(* IEC 61131-3 sources: daoli-st-library/DL_Motion (part 19) *)

(* ---- FB_DL_StringCutAlign.st ---- *)
(*==============================================================================
 * 组件名称 (Component)  : FB_DL_StringCutAlign
 * 所属子库 (Sublibrary) : DL_Motion
 * 当前版本 (Version)    : 1.0.0
 * 兼容性 (Platform)     : CODESYS 3.5 / TwinCAT 3 / 汇川 InoProShop / Machine Expert
 *                         仅依赖纯 IEC 61131-3 标准元素，零厂商方言
 * 功能描述 (Function)   : 串焊裁切对位：bCutCycle 上升沿锁存相机偏差 → 委托
 *                         FB_DL_LowPassFilter 滤波 → 比例修正计算 → 行程钳位
 *                         → 下发修正指令 → 等 bAxisInPos → 对位完成；在位等待
 *                         超时（tInPosMax，默认 T#2S）→ 中止报错（Splicer 教训
 *                         迁移：超时引脚必须带单位与默认值）。
 * 溯源 (Origin)         : 道莅 clean-room 防御性实现
 * 本文件内含 (Contains) : TYPE E_DL_AlignState / TYPE E_DL_AlignErr /
 *                         FUNCTION_BLOCK FB_DL_StringCutAlign
 * 依赖 (Depends)        : DL_Algo/FB_DL_LowPassFilter
 * 红线自检 (Redline)    : 无外部全局变量、无硬件地址直引 ｜ 全变量中英双语同行注释
 *                         防除零 + 增益/偏差钳位 + 非有限值防御 ｜ 枚举成员全部显式赋值
 *                         TON/R_TRIG/滤波器实例每周期无条件调用（仅输入条件化）｜
 *                         对位状态机 CASE 含 ELSE 兜底
 * 错误码表 (Codes)      : 16#0004_031D 就绪
 *                         16#0004_031E 信息级 偏差越界(已钳制)
 *                         16#0004_031F 信息级 修正指令已下发
 *                         16#0004_0320 故障级 在位超时(已中止)
 *                         16#0004_0321 对位完成
 * 修订历史 (Revision)   : 2026-11-17  v1.0.0  首版入库 · R27 · 阶段三批 3
 * 验收向量 (Acceptance) : 偏差 2.0 mm 增益 80% → 指令 1.6 mm；偏差 60 → 钳 50 且
 *                         031E；指令下发后 tInPosMax 内未在位 → 0320 中止
 *============================================================================*)

(*-----------------------------------------------------------------------------
 * 枚举: E_DL_AlignState（归属 DL_Motion，对位状态机状态）
 *----------------------------------------------------------------------------*)
TYPE E_DL_AlignState :
(
    eIdle    := 0,    // 就绪待节拍 / Idle, waiting for the cut cycle
    eCalc    := 10,   // 计算相：滤波 + 比例 + 钳位，下发指令 / Calculating and issuing the correction
    eWaitPos := 20,   // 等待在位相（双退出：在位成功 / 超时中止）/ Waiting for in-position, dual exit
    eDone    := 30,   // 对位完成（保持至下一节拍）/ Alignment done, held until next cycle
    eFault   := 99    // 故障兜底态 / Fault fallback
);
END_TYPE

(*-----------------------------------------------------------------------------
 * 枚举: E_DL_AlignErr（归属 DL_Motion，与 FB_DL_StringCutAlign 同文件）
 *----------------------------------------------------------------------------*)
TYPE E_DL_AlignErr :
(
    eReady    := 16#0004_031D,   // 就绪 / Ready
    eOffClamp := 16#0004_031E,   // 信息级：偏差越界已钳制 / Info: offset clamped
    eCmdSent  := 16#0004_031F,   // 信息级：修正指令已下发 / Info: correction issued
    eInPosTmo := 16#0004_0320,   // 故障级：在位超时已中止 / Fault: in-position timeout, aborted
    eAligned  := 16#0004_0321    // 对位完成 / Alignment completed
);
END_TYPE

(*==============================================================================
 * 功能块: FB_DL_StringCutAlign
 * 调用约定: 每个扫描周期无条件调用一次；tSampleTime 注入真实任务间隔。
 *============================================================================*)
FUNCTION_BLOCK FB_DL_StringCutAlign
VAR_INPUT
    fCamOffset_mm : REAL;              // 相机偏差 [毫米]，有效域 -50~50 / Camera offset [mm]
    fGainPct      : REAL := 80.0;      // 比例增益 [百分数]，有效域 0~100 / Proportional gain [percent]
    fMaxCorr_mm   : REAL := 10.0;      // 最大修正 [毫米]，须 > 0 / Maximum correction [mm]
    bCutCycle     : BOOL;              // 切割节拍触发（上升沿）/ Cut cycle trigger, rising edge
    bAxisInPos    : BOOL;              // 轴在位反馈 / Axis in-position feedback
    tInPosMax     : TIME := T#2S;      // 在位等待超时 [毫秒]，默认 T#2S / In-position timeout [ms]
    tSampleTime   : TIME := T#100MS;   // 采样周期（滤波器透传）/ Sample period, filter pass-through
END_VAR
VAR_OUTPUT
    fCorrCmd_mm   : REAL;              // 修正指令 [毫米] / Correction command [mm]
    bCorrDone     : BOOL;              // 修正完成（单拍脉冲）/ Correction done, single-scan pulse
    eErr          : E_DL_AlignErr;     // 错误码 / Error code
    eState        : E_DL_AlignState;   // 对位状态机当前状态 / Alignment state
END_VAR
VAR
    fbCutTrig     : R_TRIG;            // 切割节拍上升沿实例（无条件调用）/ Cut cycle edge instance
    fbTonInPos    : TON;               // 在位等待超时定时器（无条件调用）/ In-position timeout timer
    fbLpf         : FB_DL_LowPassFilter;   // 委托低通滤波器实例（无条件调用）/ Delegate low-pass filter instance
    fOffLatch     : REAL;              // 锁存偏差（节拍沿采样）[毫米] / Latched offset [mm]
    fOffUse       : REAL;              // 生效偏差（钳位后）[毫米] / Effective offset [mm]
    fGainUse      : REAL;              // 生效增益（钳位后）[百分数] / Effective gain [percent]
    fCorrCalc     : REAL;              // 修正计算值 [毫米] / Calculated correction [mm]
    bNonFin       : BOOL;              // 非有限输入汇总标志 / Non-finite input aggregate flag
END_VAR
VAR CONSTANT
    DL_ALN_OFF_MIN   : REAL := -50.0;   // 偏差域下限 [毫米] / Offset lower bound [mm]
    DL_ALN_OFF_MAX   : REAL := 50.0;    // 偏差域上限 [毫米] / Offset upper bound [mm]
    DL_ALN_GAIN_MIN  : REAL := 0.0;     // 增益下限 [百分数] / Gain lower bound [percent]
    DL_ALN_GAIN_MAX  : REAL := 100.0;   // 增益上限 [百分数] / Gain upper bound [percent]
    DL_ALN_INF_MAX   : REAL := 1.0E30;  // 非有限值判定幅值上限 / Magnitude bound for finite-value check
    DL_ALN_ZERO      : REAL := 0.0;     // 零值常量，避免裸字面量 / Zero constant
    DL_ALN_PCT       : REAL := 100.0;   // 百分数系数 [百分数] / Percent factor
    DL_ALN_LPF_TC    : TIME := T#100MS; // 委托滤波时间常数 [毫秒] / Delegate filter time constant [ms]
END_VAR

(*------------------------------------------------------------------------------
 * 段 1｜沿检测/TON/滤波器实例每周期无条件调用（仅输入条件化）
 *----------------------------------------------------------------------------*)
fbCutTrig(CLK := bCutCycle);                          // 节拍沿检测无条件刷新 / cycle edge refreshed unconditionally
fbTonInPos(IN := (eState = E_DL_AlignState.eWaitPos), PT := tInPosMax);   // 在位超时计时 / in-position timeout timing
fbLpf(bEnable := (eState = E_DL_AlignState.eCalc),    // 滤波仅在计算相使能 / filter enabled only in calc phase
      fIn := fOffLatch,                               // 滤波输入为锁存偏差 / filter input is the latched offset
      tTimeConst := DL_ALN_LPF_TC,                    // 滤波时间常数 [毫秒] / filter time constant [ms]
      tSampleTime := tSampleTime,                     // 采样周期透传 / sample period passed
      fOut => fOffUse);                               // 滤波输出作为生效偏差 / filtered output as effective offset

(*------------------------------------------------------------------------------
 * 段 2｜非有限值闸：偏差/增益/限幅 NaN 或溢出 → 进故障兜底态（指令撤）
 *----------------------------------------------------------------------------*)
bNonFin := (fCamOffset_mm <> fCamOffset_mm) OR (ABS(fCamOffset_mm) > DL_ALN_INF_MAX)
        OR (fGainPct      <> fGainPct)      OR (ABS(fGainPct)      > DL_ALN_INF_MAX)
        OR (fMaxCorr_mm   <> fMaxCorr_mm)   OR (ABS(fMaxCorr_mm)   > DL_ALN_INF_MAX);
IF bNonFin THEN
    eState := E_DL_AlignState.eFault;                // 进故障兜底态 / enter fault fallback
    eErr := E_DL_AlignErr.eInPosTmo;                 // 兜底并入超时段（反证句：输出同为指令撤+故障级）/ fallback mapped to timeout band
    fCorrCmd_mm := DL_ALN_ZERO;                      // 指令撤（安全侧）/ command dropped, safe side
    bCorrDone := FALSE;                              // 完成撤 / done dropped
    RETURN;
END_IF

(*------------------------------------------------------------------------------
 * 段 3｜增益与限幅参数钳位
 *----------------------------------------------------------------------------*)
fGainUse := fGainPct;                                 // 增益工作副本 / gain working copy
IF fGainUse < DL_ALN_GAIN_MIN THEN
    fGainUse := DL_ALN_GAIN_MIN;                     // 增益下限钳位 / gain floored
ELSIF fGainUse > DL_ALN_GAIN_MAX THEN
    fGainUse := DL_ALN_GAIN_MAX;                     // 增益上限钳位 / gain capped
END_IF
IF fMaxCorr_mm <= DL_ALN_ZERO THEN
    fMaxCorr_mm := 10.0;                             // 限幅非法按默认 10 mm 兜底（配置防御）/ illegal clamp falls back
END_IF

(*------------------------------------------------------------------------------
 * 段 4｜节拍沿锁存与偏差钳位（信息级 031E）
 *----------------------------------------------------------------------------*)
eErr := E_DL_AlignErr.eReady;                         // 默认就绪 / default ready
bCorrDone := FALSE;                                   // 完成脉冲逐拍先清 / done pulse cleared first
IF fbCutTrig.Q THEN
    fOffLatch := fCamOffset_mm;                       // 节拍沿锁存偏差 / latch offset on edge
    fCorrCmd_mm := DL_ALN_ZERO;                       // 新节拍指令预清 / command pre-cleared
    eState := E_DL_AlignState.eCalc;                  // 进计算相 / enter calc phase
END_IF
IF (fOffLatch < DL_ALN_OFF_MIN) OR (fOffLatch > DL_ALN_OFF_MAX) THEN
    IF fOffLatch < DL_ALN_OFF_MIN THEN
        fOffLatch := DL_ALN_OFF_MIN;                  // 偏差下限钳位 / offset floored
    ELSE
        fOffLatch := DL_ALN_OFF_MAX;                  // 偏差上限钳位 / offset capped
    END_IF
    eErr := E_DL_AlignErr.eOffClamp;                  // 信息级：偏差越界已钳制 / info: offset clamped
END_IF

(*------------------------------------------------------------------------------
 * 段 5｜对位状态机：CASE 含 ELSE 兜底
 *----------------------------------------------------------------------------*)
CASE eState OF

    E_DL_AlignState.eIdle:
        fCorrCmd_mm := DL_ALN_ZERO;                   // 就绪态指令撤 / command dropped in idle
        IF eErr = E_DL_AlignErr.eReady THEN
            eErr := E_DL_AlignErr.eReady;             // 保持就绪码 / keep ready code
        END_IF

    E_DL_AlignState.eCalc:
        fCorrCalc := fOffUse * fGainUse / DL_ALN_PCT;   // 比例修正计算 [毫米] / proportional correction [mm]
        IF fCorrCalc > fMaxCorr_mm THEN
            fCorrCalc := fMaxCorr_mm;                 // 行程上限钳位 / stroke capped
        ELSIF fCorrCalc < -fMaxCorr_mm THEN
            fCorrCalc := -fMaxCorr_mm;                // 行程下限钳位 / stroke floored
        END_IF
        fCorrCmd_mm := fCorrCalc;                     // 指令下发 [毫米] / command issued [mm]
        eErr := E_DL_AlignErr.eCmdSent;               // 信息级：指令已下发 / info: command issued
        eState := E_DL_AlignState.eWaitPos;           // 进等待在位相 / enter wait phase

    E_DL_AlignState.eWaitPos:
        IF bAxisInPos THEN
            bCorrDone := TRUE;                        // 在位成功：完成单拍脉冲 / in position: single-scan done pulse
            eErr := E_DL_AlignErr.eAligned;           // 对位完成码 / aligned code
            eState := E_DL_AlignState.eDone;          // 进完成相 / enter done phase
        ELSIF fbTonInPos.Q THEN
            eState := E_DL_AlignState.eFault;         // 在位超时：中止进故障态 / timeout: abort to fault
            eErr := E_DL_AlignErr.eInPosTmo;          // 故障级：在位超时 / fault: timeout
            fCorrCmd_mm := DL_ALN_ZERO;               // 中止撤指令（安全侧）/ abort drops command
        ELSE
            eErr := E_DL_AlignErr.eCmdSent;           // 等待中保持指令已下发码 / keep issued code while waiting
        END_IF

    E_DL_AlignState.eDone:
        fCorrCmd_mm := fCorrCalc;                     // 完成相保持指令显示 / hold command display
        IF fbCutTrig.Q THEN
            eErr := E_DL_AlignErr.eReady;             // 新节拍沿已由段 4 处理 / new edge handled in section 4
        END_IF

    E_DL_AlignState.eFault:
        fCorrCmd_mm := DL_ALN_ZERO;                   // 故障态指令撤 / command dropped in fault
        bCorrDone := FALSE;                           // 故障态完成撤 / done dropped in fault
        IF fbCutTrig.Q THEN
            eState := E_DL_AlignState.eCalc;          // 新节拍允许重试 / new cycle allows retry
        END_IF

    ELSE
        eState := E_DL_AlignState.eFault;             // 非法状态兜底 / illegal-state fallback
        eErr := E_DL_AlignErr.eInPosTmo;              // 兜底码（超时段，反证句：输出同为指令撤+故障级）/ fallback code
        fCorrCmd_mm := DL_ALN_ZERO;                   // 指令撤 / command dropped

END_CASE
END_FUNCTION_BLOCK

(* ---- FB_DL_ToolLifeBudget.st ---- *)
(*
  ==================================================================
  组件名 Component  : FB_DL_ToolLifeBudget
  分类   Category   : DL_Motion
  复杂度 Complexity  : 中
  版本   Version    : 1.0.0
  功能   Purpose    : 刀具寿命预算。切削时长（bCutting 期按 fDtSec 累计）与
                      件数（bPieceDone 沿计数）双口径累计；寿命分档预警
                      eTier：eOk / eWarn（≥fWarnPct%）/ eAlert（≥fAlertPct%）
                      / eExhausted（≥100%，置 bChangeDue）；换刀沿全量复位。
                      GitHub topics 公开语义 clean-room，与
                      FB_DL_AxisLubeDistTrig 分工。
  来源   Source     : T1-8-github-topics（刀具寿命公开语义）
  溯源   Origin     : 切削时长与件数双口径寿命预算为公开工程语义，clean-room
                      自研实现，未复制任何厂商私有库源码。
  平台   Platform   : 纯 IEC 61131-3，CODESYS / TwinCAT / InoProShop 通用
  分工声明 Split     : 与 FB_DL_AxisLubeDistTrig 分工——后者做润滑距离触发，
                      本件做刀具寿命双口径预算。
  作者   Author     : 道莅代码库 · PLC 编程专家（R59）
  ------------------------------------------------------------------
  边界 Boundary     :
                      一 非有限/组态闸：fDtSec 非有限或 ∉ (0,1] 置 bBad
                         （纪律②），冻结累计不推进（不静默吞）；
                      二 累计上界钳制（时长 1E7 秒 / 件数 1E6 件，防回绕）；
                      三 换刀沿（bToolChange 上升沿）全量复位：时长 / 件数
                         / 分档全清（解除路径唯一，R188）；
                      四 分档双口径取 max（时长比与件数比孰高），分档单调
                         不回落（锁存口径：已达档位不因当拍口径回落而降档）；
                      五 无全局变量、无外部变量声明、无物理地址寻址。
  修订记录 Revision  :
    2026-11-21  v1.0.0  R59 首版（批 4 · 序号 19）
  ==================================================================
*)

TYPE E_DL_TltTier :
(
    eTltOk       := 0,  // 寿命充足档 [-] / the healthy tier
    eTltWarn     := 10, // 预警档（≥fWarnPct%）[-] / the warn tier
    eTltAlert    := 20, // 告警档（≥fAlertPct%）[-] / the alert tier
    eTltExhausted:= 30  // 寿命耗尽档（≥100%，bChangeDue）[-] / the exhausted tier
);
END_TYPE

FUNCTION_BLOCK FB_DL_ToolLifeBudget
VAR_INPUT
    bCutting    : BOOL  := FALSE;   // 切削进行信号（时长累计闸）[-] / the cutting active signal, the time accumulation gate
    bPieceDone  : BOOL  := FALSE;   // 单件完成信号，上升沿计数 [-] / the piece done signal, the rising edge counts
    fDtSec      : LREAL := 0.1;     // 调用周期 [秒]，域 (0,1] / the call period [second]
    fLifeTimeSec: LREAL := 3600.0;  // 时长口径寿命预算 [秒] / the time budget [second]
    nLifePcs    : UDINT := 1000;    // 件数口径寿命预算 [件] / the piece budget
    fWarnPct    : LREAL := 80.0;    // 预警档阈值 [%] / the warn tier threshold [percent]
    fAlertPct   : LREAL := 95.0;    // 告警档阈值 [%] / the alert tier threshold [percent]
    bToolChange : BOOL  := FALSE;   // 换刀信号，上升沿全量复位 [-] / the tool change signal, the rising edge resets all
END_VAR
VAR_OUTPUT
    fCutTimeAcc : LREAL := 0.0;   // 切削时长累计 [秒] / the cutting time accumulated [second]
    nPieceCnt   : UDINT := 0;     // 完成件数累计 [件] / the piece count accumulated
    eTier       : E_DL_TltTier := E_DL_TltTier.eTltOk; // 寿命分档输出 [-] / the life tier outlet
    bChangeDue  : BOOL  := FALSE; // 换刀到期指示（eTltExhausted 同源）[-] / the change due indicator
    fLifePct    : LREAL := 0.0;   // 双口径寿命占用率（孰高）[%] / the life usage, the higher of the two ratios [percent]
    bBad        : BOOL  := FALSE; // 步长非有限/越域实时标志 [-] / the period fault live flag
END_VAR
VAR CONSTANT
    DL_TLT_TMAX  : LREAL := 1.0E7;  // 时长累计上界 [秒] / the time accumulation ceiling
    DL_TLT_NMAX  : UDINT := 1000000; // 件数累计上界 [件] / the piece accumulation ceiling
    DL_TLT_EPS   : LREAL := 1.0E-9; // 预算下阈值 [秒 / 件] / the budget threshold
END_VAR
VAR
    _fRatioT : LREAL; // 时长口径占用率 [%] / the time ratio [percent]
    _fRatioP : LREAL; // 件数口径占用率 [%] / the piece ratio [percent]
    _eTier   : E_DL_TltTier := E_DL_TltTier.eTltOk; // 分档锁存寄存（单调不回落）/ the tier latch, monotonic
    rtDone   : R_TRIG; // 件完成沿，段 0 无条件刷新 / the piece done edge
    rtChange : R_TRIG; // 换刀沿，段 0 无条件刷新 / the change edge
    bFinDt   : BOOL;   // 步长有限工作量 [-] / the period finiteness work flag
    bCfg     : BOOL;   // 组态域工作量 [-] / the config domain work flag
END_VAR

// 段 0｜沿检测无条件周期刷新（禁入分支，R7）/ segment 0, the unconditional refresh
rtDone(CLK := bPieceDone); // 件完成沿 / the piece done edge
rtChange(CLK := bToolChange); // 换刀沿 / the change edge

// 段 1｜换刀沿全量复位（边界三，解除路径 = 换刀沿，R188）/ segment 1, the change edge full reset
IF rtChange.Q THEN // 换刀沿 / the change edge
    fCutTimeAcc := 0.0; // 时长清零 / clear the time
    nPieceCnt := 0; // 件数清零 / clear the pieces
    _eTier := E_DL_TltTier.eTltOk; // 分档归位 / reset the tier
END_IF

// 段 2｜步长闸（边界一，实时标志非锁存）/ segment 2, the period gate
bFinDt := (fDtSec = fDtSec) AND ((fDtSec - fDtSec) = (fDtSec - fDtSec)); // 步长有限双判据（R79）/ the finiteness dual verdicts
bCfg := (fDtSec > 0.0) AND (fDtSec <= 1.0) // 步长域 (0,1] / the period domain
    AND (fLifeTimeSec > DL_TLT_EPS) AND (nLifePcs > 0) // 双口径预算为正 / the budgets positive
    AND (fWarnPct > 0.0) AND (fAlertPct > fWarnPct) AND (fAlertPct <= 100.0); // 分档阈值序合理 / the threshold order sane
bBad := (NOT bFinDt) OR (NOT bCfg); // 闸实时标志（R191 名实双出口）/ the gate flag

// 段 3｜双口径累计（闸通过才推进，上界钳制，边界一二）/ segment 3, the dual accumulation
IF bCutting AND (NOT bBad) THEN // 切削且闸通过 / cutting and gated
    fCutTimeAcc := fCutTimeAcc + fDtSec; // 时长累计 / accumulate the time
    IF fCutTimeAcc > DL_TLT_TMAX THEN // 时长上界钳制 / clamp the time ceiling
        fCutTimeAcc := DL_TLT_TMAX; // 夹到上界 / clamp
    END_IF
END_IF
IF rtDone.Q AND (NOT bBad) THEN // 件完成沿且闸通过 / the done edge and gated
    IF nPieceCnt < DL_TLT_NMAX THEN // 件数上界钳制（防回绕）/ the piece wrap guard
        nPieceCnt := nPieceCnt + 1; // 件数推进 / advance the pieces
    END_IF
END_IF

// 段 4｜分档判定（双口径孰高 + 单调锁存，边界四）/ segment 4, the tier verdict
IF (NOT bBad) AND (fLifeTimeSec > DL_TLT_EPS) AND (nLifePcs > 0) THEN // 有效预算才判定 / the verdict with the valid budgets
    _fRatioT := (fCutTimeAcc / fLifeTimeSec) * 100.0; // 时长占用率 [%]（除子域闸保证）/ the time ratio
    _fRatioP := (UDINT_TO_LREAL(nPieceCnt) / UDINT_TO_LREAL(nLifePcs)) * 100.0; // 件数占用率 [%]/ the piece ratio
    IF _fRatioT > _fRatioP THEN // 孰高口径 / the higher ratio
        fLifePct := _fRatioT; // 取时长口径 / take the time ratio
    ELSE // 件数口径更高或持平 / the piece ratio higher or equal
        fLifePct := _fRatioP; // 取件数口径 / take the piece ratio
    END_IF
    IF fLifePct >= 100.0 THEN // 耗尽档 / the exhausted tier
        _eTier := E_DL_TltTier.eTltExhausted; // 升档（锁存单调）/ raise the tier
    ELSIF fLifePct >= fAlertPct THEN // 告警档 / the alert tier
        IF _eTier < E_DL_TltTier.eTltAlert THEN // 仅低档升档（单调不回落）/ raise only from a lower tier
            _eTier := E_DL_TltTier.eTltAlert; // 升到告警 / raise to the alert
        END_IF
    ELSIF fLifePct >= fWarnPct THEN // 预警档 / the warn tier
        IF _eTier < E_DL_TltTier.eTltWarn THEN // 仅低档升档 / raise only from a lower tier
            _eTier := E_DL_TltTier.eTltWarn; // 升到预警 / raise to the warn
        END_IF
    END_IF
END_IF
eTier := _eTier; // 分档出口 / the tier outlet
bChangeDue := (_eTier = E_DL_TltTier.eTltExhausted); // 换刀到期（R191 名实双出口）/ the change due indicator
END_FUNCTION_BLOCK

(* ---- FB_DL_TrackerAngleYearWin.st ---- *)
(*
  FB_DL_TrackerAngleYearWin  —  跟踪支架年度角度表切换 / Tracker annual angle-table switching
  分类 Category : DL_Motion
  码位 Code     : 16#04_0_A1
  版本 Version  : 1.0.0
  溯源 Source   : LGF DateAndTimer 语义借鉴 · clean-room 实现，仅借分类/参数域/命名，未复制源码
  功能 Function : 1) 年窗 + 月窗双闸同时生效才允许角度表切换（任一窗不开即禁止）；
                  2) 角度表切换仅在「双窗生效 + 支架静止」时执行；运动中切换排队到停止（bSwitchPending）；
                  3) 表版本号锁存，切换瞬间只给出新版本号单点，防半新半旧。
  边界 Boundary : ① 年窗/月窗参数越界钳位照算（报码不拒算）；
                  ② 仅在「双窗同时生效 + 支架静止」执行切换，运动中排队到停止；
                  ③ 表版本锁存防切换瞬间半新半旧；
                  ④ 输出三行同向：双窗标志 → 版本号 → 切换待决标志。
  依赖 Depends  : FB_DL_YearWindowCheck、FB_DL_MonthWindowCheck（均每拍无条件调用）

  码表 Error codes（本件子码步进 16#10，避让邻件码位）:
    16#0002_04A1 故障级：年窗组态非法（空窗/日期越界钳位后仍非法）
    16#0002_04B1 故障级：月窗组态非法（目标日为 0 或窗宽越界）
    16#0002_04C1 信息级：日期注入越界已钳位照算 / 运动中的切换排队（不置 bError）
*)

TYPE E_DL_TayPhase :
(
    eIdle    := 0,   // 空闲 / Idle
    eWait    := 10,  // 等双窗与静止 / Waiting for both windows and standstill
    ePending := 20,  // 切换排队中 / Switch pending
    eSwitch  := 30,  // 执行切换 / Switching
    eFault   := 90   // 组态故障锁定 / Configuration fault locked
);
END_TYPE

FUNCTION_BLOCK FB_DL_TrackerAngleYearWin
VAR_INPUT
    bEnable       : BOOL;                          // 总使能，FALSE 回空闲 / Master enable
    bReset        : BOOL;                          // 复位，上升沿清组态故障 / Reset, clears configuration fault
    nYear         : INT := 2026;                   // 当前年 [年]，域 1970~2099 / Current year [year]
    nMonth        : INT := 1;                      // 当前月 [月]，域 1~12 / Current month [month]
    nDay          : INT := 1;                      // 当前日 [日]，域 1~31 / Current day [day]
    nStartYear    : INT := 2026;                   // 年窗起始年 [年] / Window start year [year]
    nStartMonth   : INT := 1;                      // 年窗起始月 [月] / Window start month [month]
    nStartDay     : INT := 1;                       // 年窗起始日 [日] / Window start day [day]
    nEndYear      : INT := 2026;                   // 年窗结束年 [年] / Window end year [year]
    nEndMonth     : INT := 12;                     // 年窗结束月 [月] / Window end month [month]
    nEndDay       : INT := 31;                     // 年窗结束日 [日] / Window end day [day]
    nTargetDay    : INT := 15;                     // 月窗目标日（正 = 第 N 天，负 = 月末倒数）[日] / Month target day
    nWindowDays   : INT := 3;                      // 月窗宽度 [日]，域 1~31 / Month window width [days]
    nYearMonth    : INT := 3;                      // 年度窗生效月份 [月]，域 1~12 / Yearly month [month]
    bTrackerStill : BOOL;                          // 支架静止标志（速度为 0 且无运动命令）/ Tracker standstill flag
    nTableVerNew  : INT := 2;                      // 新角度表版本号 [版本]，域 >= 1 / New angle table version
    nTableVerCur  : INT := 1;                      // 当前生效版本号 [版本]，域 >= 1 / Current active version
END_VAR
VAR_OUTPUT
    bYearWin      : BOOL;                          // 年窗生效 / Year window active
    bMonthWin     : BOOL;                          // 月窗生效 / Month window active
    bBothWin      : BOOL;                          // 双窗同时生效 / Both windows active
    nTableVerLatched : INT;                        // 锁存并生效的表版本号 [版本] / Latched table version
    bSwitchPending: BOOL;                          // 切换排队中（运动中）/ Switch pending during motion
    bSwitched     : BOOL;                          // 切换完成（单拍脉冲）/ Switch completed, single pulse
    bError        : BOOL;                          // 故障标志，与故障级码配对 / Fault flag paired with fault codes
    uErrorId      : UDINT;                         // 事件码，0 = 无事件 / Event code, 0 = none
    eStateOut     : E_DL_TayPhase;                 // 状态机当前态，段尾单点映射 / Phase mapped at tail
END_VAR
VAR
    _eState       : E_DL_TayPhase := E_DL_TayPhase.eIdle;  // 内部状态 / Internal state
    rtrReset      : R_TRIG;                        // 复位沿 / Reset edge
    fbYearWin     : FB_DL_YearWindowCheck;         // 年窗实例（无条件调用）/ Year window instance
    fbMonthWin    : FB_DL_MonthWindowCheck;        // 月窗实例（无条件调用）/ Month window instance
    nYearC        : INT;                           // 钳位后当前年 [年] / Clamped current year
    nMonthC       : INT;                           // 钳位后当前月 [月] / Clamped current month
    nDayC         : INT;                           // 钳位后当前日 [日] / Clamped current day
    bYWin         : BOOL;                          // 年窗结果暂存 / Year window buffer
    bMWin         : BOOL;                          // 月窗结果暂存 / Month window buffer
    uFault        : UDINT;                         // 锁存故障码 / Latched fault code
    uInfo         : UDINT;                         // 信息级码 / Information code
END_VAR
VAR CONSTANT
    DL_TAY_YMIN   : INT := 1970;                   // 年份物理域下限 [年] / Year domain low
    DL_TAY_YMAX   : INT := 2099;                   // 年份物理域上限 [年] / Year domain high
    DL_TAY_DMAX   : INT := 31;                     // 日物理域上限 [日] / Day domain high
END_VAR

(* === 段 0 · 实例刷新（无条件周期调用）=== *)
rtrReset(CLK := bReset);                          // 每拍刷新复位沿

(* === 段 1 · 参数钳位（越界钳定照算，报码不拒算）=== *)
nYearC := nYear;                                  // 年份钳位
IF nYearC < DL_TAY_YMIN THEN
    nYearC := DL_TAY_YMIN;
END_IF
IF nYearC > DL_TAY_YMAX THEN
    nYearC := DL_TAY_YMAX;
END_IF
nMonthC := nMonth;                                // 月份钳位
IF nMonthC < 1 THEN
    nMonthC := 1;
END_IF
IF nMonthC > 12 THEN
    nMonthC := 12;
END_IF
nDayC := nDay;                                    // 日期钳位
IF nDayC < 1 THEN
    nDayC := 1;
END_IF
IF nDayC > DL_TAY_DMAX THEN
    nDayC := DL_TAY_DMAX;
END_IF
uInfo := 16#0000;                                 // 信息码每拍清零
IF (nYear <> nYearC) OR (nMonth <> nMonthC) OR (nDay <> nDayC) THEN
    uInfo := 16#0002_04C1;                        // 信息级：日期注入越界已钳位照算
END_IF

(* === 段 2 · 年窗实例（每拍无条件调用）=== *)
fbYearWin(bEnable := bEnable,
          bReset := rtrReset.Q,
          nYear := nYearC,
          nMonth := nMonthC,
          nDay := nDayC,
          nStartYear := nStartYear,
          nStartMonth := nStartMonth,
          nStartDay := nStartDay,
          nEndYear := nEndYear,
          nEndMonth := nEndMonth,
          nEndDay := nEndDay,
          bIncludeEnd := TRUE);                   // 结束日含当天（闭区间）
bYWin := fbYearWin.bInWindow;                     // 年窗结果
bYearWin := bYWin;                                // 年窗输出
IF fbYearWin.bInvalidConfig THEN
    uFault := 16#0002_04A1;                       // 故障级：年窗组态非法（空窗）
END_IF

(* === 段 3 · 月窗实例（每拍无条件调用）=== *)
fbMonthWin(bEnable := bEnable,
           nYear := INT_TO_DINT(nYearC),          // 标准转换函数
           nMonth := INT_TO_DINT(nMonthC),
           nDay := INT_TO_DINT(nDayC),
           nTargetDay := INT_TO_DINT(nTargetDay),
           nWindowDays := INT_TO_DINT(nWindowDays),
           bYearly := TRUE,                       // 年度窗：仅生效月份开放
           nYearMonth := INT_TO_DINT(nYearMonth));
bMWin := fbMonthWin.bInWindow;                    // 月窗结果
bMonthWin := bMWin;                               // 月窗输出
IF (nTargetDay = 0) OR (nWindowDays < 1) OR (nWindowDays > DL_TAY_DMAX)
   OR (nYearMonth < 1) OR (nYearMonth > 12) THEN
    uFault := 16#0002_04B1;                       // 故障级：月窗组态非法
END_IF
IF rtrReset.Q THEN
    uFault := 16#0000;                            // 复位沿清锁存（复位路径可达）
    bSwitched := FALSE;                           // 切换脉冲复位（非置位型）
END_IF
bBothWin := bYWin AND bMWin;                      // 双窗同时生效

(* === 段 4 · 主状态机（ENUM + CASE，含 ELSE 兜底）=== *)
CASE _eState OF
E_DL_TayPhase.eIdle :
    bSwitched := FALSE;                           // 空闲无切换脉冲
    bSwitchPending := FALSE;                      // 无排队
    IF uFault <> 16#0000 THEN
        _eState := E_DL_TayPhase.eFault;          // 组态故障优先
    ELSIF bEnable THEN
        _eState := E_DL_TayPhase.eWait;           // 进入等待相
    END_IF

E_DL_TayPhase.eWait :
    IF NOT bBothWin THEN
        bSwitchPending := FALSE;                  // 双窗不满足：排队取消
    ELSIF bBothWin AND (NOT bTrackerStill) THEN
        bSwitchPending := TRUE;                   // 运动中：排队到停止
        uInfo := 16#0002_04C1;                    // 信息级：运动中的切换排队
        _eState := E_DL_TayPhase.ePending;
    ELSIF bBothWin AND bTrackerStill AND (nTableVerNew <> nTableVerCur) THEN
        _eState := E_DL_TayPhase.eSwitch;         // 双窗 + 静止 + 版本不同：执行切换
    ELSE
        nTableVerLatched := nTableVerCur;         // 版本一致：锁存当前版本
    END_IF

E_DL_TayPhase.ePending :
    bSwitchPending := TRUE;                       // 排队标志保持
    IF NOT bBothWin THEN
        bSwitchPending := FALSE;                  // 窗关闭：排队取消
        _eState := E_DL_TayPhase.eWait;
    ELSIF bTrackerStill THEN
        bSwitchPending := FALSE;                  // 支架静止：排队结束（可到达的解除路径）
        _eState := E_DL_TayPhase.eSwitch;         // 转执行切换
    END_IF

E_DL_TayPhase.eSwitch :
    IF bTrackerStill AND bBothWin THEN
        nTableVerLatched := nTableVerNew;         // 单点锁存新版本（防半新半旧）
        bSwitched := TRUE;                        // 置位型：切换完成脉冲（段尾不清零）
        _eState := E_DL_TayPhase.eWait;           // 回等待相
    ELSIF NOT bTrackerStill THEN
        bSwitchPending := TRUE;                   // 运动中：回排队（不切换）
        _eState := E_DL_TayPhase.ePending;
    ELSIF NOT bBothWin THEN
        _eState := E_DL_TayPhase.eWait;           // 窗关闭：放弃切换
    END_IF

E_DL_TayPhase.eFault :
    bSwitchPending := FALSE;                      // 故障态取消排队
    nTableVerLatched := nTableVerCur;             // 版本保持当前（不切表）
    IF uFault = 16#0000 THEN
        _eState := E_DL_TayPhase.eIdle;           // 解锁回空闲
    END_IF

ELSE
    _eState := E_DL_TayPhase.eFault;              // 非法状态拦截
    uFault := 16#0002_04A1;                       // 故障级：相 ID 越界
    nTableVerLatched := nTableVerCur;             // 安全侧保持当前版本
    bSwitched := FALSE;                           // 安全侧不报切换
END_CASE
IF NOT bEnable THEN
    _eState := E_DL_TayPhase.eIdle;               // 失能最高优先回空闲
    bSwitchPending := FALSE;                      // 取消排队
    bSwitched := FALSE;                           // 切换脉冲复位
END_IF

(* === 段 5 · 输出映射（三行同向：双窗 → 版本号 → 排队标志）=== *)
IF nTableVerLatched < 1 THEN
    nTableVerLatched := nTableVerCur;             // 版本号非法兜底：保持当前（防 0 版本）
END_IF
bError := (uFault <> 16#0000);                    // 故障标志仅由故障级码置位（R45 配对）
IF bError THEN
    uErrorId := uFault;                           // 故障级优先上报
ELSE
    uErrorId := uInfo;                            // 否则上报信息级码
END_IF
eStateOut := _eState;                             // 输出枚举段尾单点映射（N2 规则）
END_FUNCTION_BLOCK

(* ---- FB_DL_TrackerBacktrackCalc.st ---- *)
// =====================================================================
// FB_DL_TrackerBacktrackCalc.st
// 光伏跟踪支架逆跟踪角度修正（阵列阴影几何, 逐排互遮挡角计算）
// PV tracker backtracking angle with array shading geometry
// 所属子库: DL_Motion    版本: v1.0.0    兼容: CODESYS V3.5+ / TwinCAT 3 / 汇川 InoProShop
// 码位: 16#0004_0354 ~ 16#0004_0358 (本件独占 5 槽, 勿复用)
// 溯源: 道莅 clean-room 防御性实现
//       来源组标签: photovoltaic, solar-tracker, backtrack, geometry
// 修改记录: R30 初版 (ROUND_PLAN_R30 序 14)
// 分层声明: 太阳高度角/方位角经引脚注入（上游消费太阳位置计算件输出）,
//           本件为逐排阴影几何层, 每拍全量重算
// 几何模型: 面板绕南北轴旋转角 R, 收集宽度 W, 排间距 P;
//           面板端点高 h = (W/2)·sin(R), 水平投影 d = (W/2)·cos(R);
//           无遮挡约束 d + h/tan(高角) ≤ P − W/2;
//           解 a·cos(R) + b·sin(R) = K（a=W/2, b=W/(2·tan(高角)), K=P−W/2）
//           得 R_limit = asin(K/√(a²+b²)) − atan(b/a), 全程 arctan/asin 防除零
// =====================================================================
FUNCTION_BLOCK FB_DL_TrackerBacktrackCalc
VAR_INPUT
    fSunElev_deg   : REAL := 30.0;  // 太阳高度角 -90~90 度（注入）/ Sun elevation [deg]
    fSunAzi_deg    : REAL := 180.0; // 太阳方位角 0~360 度（注入）/ Sun azimuth [deg]
    fRowPitch_m    : REAL := 6.0;   // 排间距 0.5~20 m / Row pitch [m]
    fCollectWidth_m: REAL := 2.0;   // 收集宽度（面板展开占宽）0~50 m / Collector width [m]
    fMaxAngle_deg  : REAL := 60.0;  // 机械限位角 0~90 度 / Mechanical limit angle [deg]
END_VAR
VAR_OUTPUT
    fTrackAngle_deg  : REAL := 0.0;   // 跟踪支架角度, 安全侧 0 度 / Track angle [deg]
    bBacktrackActive : BOOL := FALSE; // 逆跟踪激活标志 / Backtracking active flag
    fShadeLimit_deg  : REAL := 0.0;   // 阴影约束限角 0~90 度 / Shade limit angle [deg]
    eErr             : UDINT := 16#0004_0354;  // 错误码 / Error code
END_VAR
VAR
    rPi       : REAL := 3.14159265358979;   // 圆周率 / Pi constant
    bCfgErr   : BOOL := FALSE;        // 组态非法标记 / Configuration error flag
    bClampInfo: BOOL := FALSE;        // 输出限幅信息标记 / Output clamp info flag
    fElevR    : REAL := 0.0;          // 高度角弧度 / Elevation in radian [rad]
    fAziR     : REAL := 0.0;          // 方位角弧度 / Azimuth in radian [rad]
    fXew      : REAL := 0.0;          // 太阳矢量东西向投影 / Sun east-west projection
    fZup      : REAL := 0.0;          // 太阳矢量天顶向投影 / Sun up projection
    fIdealR   : REAL := 0.0;          // 理想跟踪角弧度 / Ideal track angle [rad]
    fA        : REAL := 0.0;          // 几何系数 a = W/2 / Geometry coefficient a
    fB        : REAL := 0.0;          // 几何系数 b = W/(2·tan(高角)) / Geometry coefficient b
    fK        : REAL := 0.0;          // 几何常数 K = P − W/2 / Geometry constant K
    fDen      : REAL := 0.0;          // 系数模长 / Coefficient modulus
    fRatio    : REAL := 0.0;          // 反正弦自变量 / Arcsine argument
    fPhiR     : REAL := 0.0;          // 相位角弧度 / Phase angle [rad]
    fRlimR    : REAL := 0.0;          // 阴影限角弧度 / Shade limit [rad]
    fIdealD   : REAL := 0.0;          // 理想跟踪角度 / Ideal track angle [deg]
    fLastAng  : REAL := 0.0;          // 上次有效输出角保持量 / Last valid angle hold [deg]
    xHasLast  : BOOL := FALSE;        // 已有有效输出标记 / Has valid output flag
END_VAR

// ---------------------------------------------------------------------
// 代码位表（本件独占, 勿复用）:
//   16#0004_0354 信息 跟踪角正常（未触发逆跟踪, 含太阳高度角不大于 0 时归位 0 度）
//   16#0004_0355 信息 逆跟踪激活（阴影约束生效, 限角压向跟踪输出）
//   16#0004_0356 信息 输出限幅生效（理想角越出机械限位, 信息级）
//   16#0004_0357 故障 太阳角输入非有限（保持上次有效角, 不新增动作）,
//                解除式 = 输入恢复有限
//   16#0004_0358 故障 组态非法（排间距越出 0.5~20 m, 宽度/限位角非法）,
//                解除式 = 恢复合法组态
// ---------------------------------------------------------------------

// ---- 组态闸 / Configuration gate ----
bCfgErr := FALSE;                   // 复位 / Reset
IF (fRowPitch_m <> fRowPitch_m) OR (fRowPitch_m < 0.5) OR (fRowPitch_m > 20.0) THEN
    bCfgErr := TRUE;                // 排间距非法 / Illegal row pitch
END_IF
IF (fCollectWidth_m <> fCollectWidth_m) OR (fCollectWidth_m <= 0.0) OR (fCollectWidth_m > 50.0) THEN
    bCfgErr := TRUE;                // 收集宽度非法 / Illegal width
END_IF
IF (fMaxAngle_deg <> fMaxAngle_deg) OR (fMaxAngle_deg <= 0.0) OR (fMaxAngle_deg > 90.0) THEN
    bCfgErr := TRUE;                // 限位角非法 / Illegal limit angle
END_IF

// ---- 输出缺省 / Output defaults ----
bBacktrackActive := FALSE;          // 缺省非逆跟踪 / Default no backtrack
bClampInfo := FALSE;                // 缺省无限幅 / Default no clamp
fShadeLimit_deg := 0.0;             // 缺省零 / Default zero

// ---- 非有限太阳角: 保持上次有效角（安全侧不新增动作）/ Non-finite sun: hold last ----
IF bCfgErr THEN
    fTrackAngle_deg := 0.0;         // 组态非法安全侧归零 / Config fault safe zero
    eErr := 16#0004_0358;           // 组态码 / Config code
ELSIF (fSunElev_deg <> fSunElev_deg) OR (ABS(fSunElev_deg) >= 1.0E12)
   OR (fSunAzi_deg <> fSunAzi_deg) OR (ABS(fSunAzi_deg) >= 1.0E12) THEN
    fTrackAngle_deg := fLastAng;    // 保持上次有效角 / Hold last valid angle
    eErr := 16#0004_0357;           // 非有限码 / Non-finite code
ELSIF fSunElev_deg <= 0.0 THEN
    // 太阳高度角不大于 0 → 归位停跟踪（安全侧 0 度）/ Night: park at 0 degree
    fTrackAngle_deg := 0.0;
    fLastAng := 0.0;                // 保持量同步归位 / Hold value parked
    xHasLast := TRUE;               // 置有效标记 / Set valid flag
    eErr := 16#0004_0354;           // 正常归位 / Normal park
ELSE
    // ---- 每拍全量重算 / Full recalculation each cycle ----
    fElevR := fSunElev_deg * rPi / 180.0;   // 高度角弧度 / Elevation radian
    fAziR  := fSunAzi_deg * rPi / 180.0;    // 方位角弧度 / Azimuth radian
    fXew   := COS(fElevR) * SIN(fAziR);     // 东西向投影 / East-west projection
    fZup   := SIN(fElevR);                  // 天顶向投影 / Up projection
    IF fZup < 0.05 THEN
        fZup := 0.05;           // 天顶分量下限防除零 / Up floor against division
    END_IF
    fIdealR := ATAN(fXew / fZup);           // 理想跟踪角弧度 / Ideal angle [rad]
    fIdealD := fIdealR * 180.0 / rPi;       // 理想角度数 / Ideal angle [deg]

    // ---- 阴影几何求限角 / Shading geometry limit ----
    IF fSunElev_deg < 1.0 THEN
        fRlimR := 0.0;          // 近地平角限角归零（贴平放） / Near horizon: flat limit
    ELSE
        fA := fCollectWidth_m * 0.5;                    // a = W/2 / Coefficient a
        fB := fA / TAN(fElevR);                         // b = W/(2·tan) / Coefficient b
        fK := fRowPitch_m - fA;                         // K = P − W/2 / Constant K
        fDen := SQRT((fA * fA) + (fB * fB));            // 模长 / Modulus
        fRatio := fK / fDen;                            // 反正弦自变量 / Arcsine argument
        IF fRatio > 1.0 THEN
            fRlimR := fMaxAngle_deg * rPi / 180.0;      // 阳光充足无阴影约束 / No shade constraint
        ELSIF fRatio < -1.0 THEN
            fRlimR := 0.0;      // 几何不可达, 限角归零 / Unreachable geometry, flat limit
        ELSE
            fPhiR  := ATAN(fB / fA);                    // 相位角（a 恒正防除零）/ Phase angle
            fRlimR := ASIN(fRatio) - fPhiR;             // 解临界角 / Solve critical angle
        END_IF
    END_IF
    // 限角归一到 0~限位 / Normalize limit to 0..max
    IF fRlimR < 0.0 THEN
        fRlimR := 0.0;          // 下界钳位 / Clamp lower
    END_IF
    IF fRlimR > (fMaxAngle_deg * rPi / 180.0) THEN
        fRlimR := fMaxAngle_deg * rPi / 180.0;      // 上界钳位 / Clamp upper
    END_IF
    fShadeLimit_deg := fRlimR * 180.0 / rPi;        // 输出限角度数 / Output limit [deg]

    // ---- 逆跟踪判定与输出 / Backtracking decision and output ----
    IF ABS(fIdealD) <= fShadeLimit_deg THEN
        fTrackAngle_deg := fIdealD;             // 未越限直接跟踪 / Track ideal
        bBacktrackActive := FALSE;              // 非逆跟踪 / Not backtracking
    ELSE
        bBacktrackActive := TRUE;               // 拍 N 进入逆跟踪 / Backtracking active
        IF fIdealD >= 0.0 THEN
            fTrackAngle_deg := fShadeLimit_deg; // 正向压到限角 / Positive side limited
        ELSE
            fTrackAngle_deg := -fShadeLimit_deg;    // 反向压到限角 / Negative side limited
        END_IF
    END_IF
    // 机械限位钳位（信息级）/ Mechanical clamp with info code
    IF fTrackAngle_deg > fMaxAngle_deg THEN
        fTrackAngle_deg := fMaxAngle_deg;       // 上限钳位 / Clamp upper
        bClampInfo := TRUE;                     // 置限幅信息 / Set clamp info
    END_IF
    IF fTrackAngle_deg < (-fMaxAngle_deg) THEN
        fTrackAngle_deg := -fMaxAngle_deg;      // 下限钳位 / Clamp lower
        bClampInfo := TRUE;
    END_IF
    fLastAng := fTrackAngle_deg;    // 更新有效保持量 / Update hold value
    xHasLast := TRUE;               // 置有效标记 / Set valid flag

    // ---- 错误码仲裁 / Error arbitration ----
    IF bClampInfo THEN
        eErr := 16#0004_0356;       // 限幅信息 / Clamp info
    ELSIF bBacktrackActive THEN
        eErr := 16#0004_0355;       // 逆跟踪信息 / Backtrack info
    ELSE
        eErr := 16#0004_0354;       // 正常 / Normal
    END_IF
END_IF

END_FUNCTION_BLOCK

(* ---- FB_DL_TrackerMotDiag.st ---- *)
// =====================================================================
// FB_DL_TrackerMotDiag.st
// 跟踪支架回转减速机健康诊断（电流偏差 + 跟随误差 EWMA → 0~100 评分）
// Tracker drive health diagnosis FB
// 码位: 16#0004_034A ~ 16#0004_034E (本件独占 5 槽)
// 修改记录: R29 初版 (按 DISPATCH_R29 序 14)
// =====================================================================
FUNCTION_BLOCK FB_DL_TrackerMotDiag
VAR_INPUT
    bEnable        : BOOL  := FALSE;   // 使能 / Enable
    bReset         : BOOL  := FALSE;   // 复位锁存 / Reset
    fCurrent_A     : REAL  := 0.0;     // 电机电流 0~200 A / Motor current [A]
    fBaseCurrent_A : REAL  := 5.0;     // 标定基线电流 >0 A / Baseline current [A]
    fFollowErr_deg : REAL  := 0.0;     // 跟随误差 -10~10 ° / Following error [deg]
    fSpeed_degS    : REAL  := 0.0;     // 转速 -5~5 °/s / Speed [deg/s]
    fSpeedMin_degS : REAL  := 0.05;    // 判定运行的最小转速 >0 °/s / Min speed [deg/s]
    fErrMax_deg    : REAL  := 1.0;     // 跟随误差报警 0.01~20 ° / Max following error [deg]
    fCurDevMax_pct : REAL  := 60.0;    // 电流偏差报警 5~300 % / Max current deviation [%]
    fAlpha         : REAL  := 0.2;     // EWMA 系数 (0,1] / EWMA factor [-]
END_VAR
VAR_OUTPUT
    fCurDev_pct    : REAL;             // 电流相对偏差 % / Current deviation [%]
    fEwmaErr_deg   : REAL;             // 跟随误差 EWMA ° / EWMA error [deg]
    uScore         : USINT;            // 健康评分 0~100 / Health score
    bWarn          : BOOL;             // 预警（评分 < 60）/ Warning
    bAlarm         : BOOL;             // 报警（评分 < 30 或越限，锁存）/ Alarm latched
    eErr           : UDINT;            // 错误码 / Error code
END_VAR
VAR
    fScoreR        : REAL;             // 评分实数中间量 / Score real intermediate [-]
    fAlphaSafe     : REAL;             // 钳位后 EWMA 系数 / Clamped alpha [-]
    bMoving        : BOOL;             // 运行判 / Moving flag
    xFirstScan     : BOOL  := TRUE;    // 首扫标记 / First-scan flag
END_VAR

// ---------------------------------------------------------------------
// 代码位表（本件独占，勿复用）:
//   16#0004_034A 信息 诊断正常（评分 ≥ 60）
//   16#0004_034B 故障 输入非有限
//   16#0004_034C 故障 fBaseCurrent_A ≤ 0 / fAlpha ≤ 0 或 >1 / fErrMax_deg ≤ 0（组态错）
//   16#0004_034D 信息 静止（ABS(fSpeed_degS) < fSpeedMin_degS）→ 电流项保持上次值，仅更误差项
//   16#0004_034E 故障 fCurDev_pct > fCurDevMax_pct 或 ABS(fEwmaErr_deg) > fErrMax_deg → bAlarm=TRUE 锁存
// ---------------------------------------------------------------------

// ---- 非有限闸 / Finite gate ----
IF (fCurrent_A <> fCurrent_A) OR (ABS(fCurrent_A) >= 1.0E12)
   OR (fBaseCurrent_A <> fBaseCurrent_A) OR (ABS(fBaseCurrent_A) >= 1.0E12)
   OR (fFollowErr_deg <> fFollowErr_deg) OR (ABS(fFollowErr_deg) >= 1.0E12)
   OR (fSpeed_degS <> fSpeed_degS) OR (ABS(fSpeed_degS) >= 1.0E12)
   OR (fSpeedMin_degS <> fSpeedMin_degS) OR (ABS(fSpeedMin_degS) >= 1.0E12)
   OR (fErrMax_deg <> fErrMax_deg) OR (ABS(fErrMax_deg) >= 1.0E12)
   OR (fCurDevMax_pct <> fCurDevMax_pct) OR (ABS(fCurDevMax_pct) >= 1.0E12)
   OR (fAlpha <> fAlpha) OR (ABS(fAlpha) >= 1.0E12) THEN
    eErr := 16#0004_034B;       // 故障码 / Fault code
    RETURN;                     // 输出保持 / Outputs hold
END_IF

// ---- 组态错闸 / Configuration fault gate ----
IF (fBaseCurrent_A <= 0.0) OR (fAlpha <= 0.0) OR (fAlpha > 1.0) OR (fErrMax_deg <= 0.0) THEN
    eErr := 16#0004_034C;       // 故障码 / Fault code
    RETURN;                     // 输出保持 / Outputs hold
END_IF

// ---- 首扫：EWMA 初值 = 当拍误差（R16 首扫纪律）/ First scan: EWMA init = current error ----
IF xFirstScan THEN
    fEwmaErr_deg := fFollowErr_deg;     // 初值 / Init
    xFirstScan := FALSE;        // 清标记 / Clear flag
END_IF

// ---- 使能撤销 / Disable ----
IF NOT bEnable THEN
    bWarn := FALSE;             // 预警复位 / Warn reset
    eErr := 16#0004_034A;       // 信息级：空闲 / Info: idle
    RETURN;                     // 评分与报警锁存保持 / Score and latch hold
END_IF

// ---- 运行判 / Moving check ----
bMoving := (ABS(fSpeed_degS) >= fSpeedMin_degS);    // 运行标志 / Moving flag

// ---- 跟随误差 EWMA（3 行内联）/ EWMA inline ----
fEwmaErr_deg := fEwmaErr_deg + fAlpha * (fFollowErr_deg - fEwmaErr_deg);    // EWMA / EWMA update

// ---- 电流偏差（分母下限闸已由组态错保证 >0）/ Current deviation ----
IF bMoving THEN
    fCurDev_pct := (fCurrent_A - fBaseCurrent_A) / fBaseCurrent_A * 100.0;  // 相对偏差 % / Deviation [%]
    IF fCurDev_pct < 0.0 THEN
        fCurDev_pct := 0.0;     // 轻载不算负偏差 / Light load not negative
    END_IF
END_IF
// 静止时电流项保持上次值（电流无意义，不误判堵转）/ Stationary: hold current term

// ---- 报警锁存（越限判 + 解除路径）/ Alarm latch with release path ----
IF bAlarm THEN
    // 锁存回放，不按当下输入重推断 / Latched replay
    eErr := 16#0004_034E;       // 故障码回放 / Fault code replay
    IF bReset
       AND (fCurDev_pct <= fCurDevMax_pct)
       AND (ABS(fEwmaErr_deg) <= fErrMax_deg) THEN
        bAlarm := FALSE;        // 解除：越限量已回落 / Release when back under limits
    END_IF
    RETURN;                     // 锁存中评分冻结 / Score frozen while latched
END_IF

// ---- 越限直接报警（堵转/异物 或 跟随误差超限）/ Direct alarm on limits ----
IF (fCurDev_pct > fCurDevMax_pct) OR (ABS(fEwmaErr_deg) > fErrMax_deg) THEN
    bAlarm := TRUE;             // 锁存 / Latch
    eErr := 16#0004_034E;       // 故障码 / Fault code
    RETURN;                     // 本拍结束 / End of cycle
END_IF

// ---- 健康评分 / Health score ----
// 公式：100 - 0.5×max(0, fCurDev_pct-20) - 20×ABS(fEwmaErr_deg)/fErrMax_deg
fScoreR := 100.0
           - 0.5 * (fCurDev_pct - 20.0)      // 电流偏差罚项（负值由判 max 处理）/ Current penalty
           - 20.0 * ABS(fEwmaErr_deg) / fErrMax_deg;     // 误差罚项 / Error penalty
IF fCurDev_pct <= 20.0 THEN
    // 电流偏差 ≤20 % 无电流罚项 / No current penalty under 20 %
    fScoreR := 100.0 - 20.0 * ABS(fEwmaErr_deg) / fErrMax_deg;  // 只含误差罚项 / Error only
END_IF
// 结果钳 [0,100] / Clamp score
IF fScoreR > 100.0 THEN
    fScoreR := 100.0;           // 上限 / Upper clamp
ELSIF fScoreR < 0.0 THEN
    fScoreR := 0.0;             // 下限 / Lower clamp
END_IF
// TRUNC 取整（禁止 TRUNC+1，R28 整数进位纪律）/ Truncate, no +1
uScore := REAL_TO_USINT(TRUNC(fScoreR));    // 评分输出 / Score output

// ---- 预警判 / Warn verdict ----
bWarn := (uScore < 60);         // 评分 < 60 预警 / Warn under 60

// ---- 错误码 / Error code ----
IF bWarn THEN
    eErr := 16#0004_034D;       // 信息级：预警或静止登记 / Info: warn or stationary
ELSE
    eErr := 16#0004_034A;       // 信息级：诊断正常 / Info: normal
END_IF

// ---- 静止信息级覆盖 / Stationary info override ----
IF NOT bMoving THEN
    eErr := 16#0004_034D;       // 信息级：静止只更误差项 / Info: stationary
END_IF

END_FUNCTION_BLOCK

(* ---- FB_DL_TrackerSnowShedAngle.st ---- *)
//==============================================================================
// 功能块：FB_DL_TrackerSnowShedAngle ｜ 中文名称：跟踪支架雪载卸荷角与复位
// 所属子库：DL_Motion ｜ 版本：v1.0.0 ｜ 兼容：CODESYS V3.5+ / TwinCAT 3 / 汇川 InoProShop
// 功能描述：雪载卸荷顺控——采暖季窗有效（bHeatSeason 电平，由上层日历
//           窗给出）且雪载超阈值 → 目标角切卸荷角（限速逼近，保护减速
//           机与雪载静摩擦）；卸荷保持最短时间后才允许退出（防雪未滑
//           落即回摆重复触发）；退出条件 = 雪载 < 阈值 - 回差 或 采暖季
//           结束，且保持最短时间已满 → 目标角切回正常跟踪角（透传输入，
//           限速逼近）。角反馈全程跟踪校验：反馈与命令偏差超容差持续
//           超窗 → 判跟踪失败，冻结命令安全侧并报故障。
// 遗留假设（R95 代理阈值三句）：① 代理值 = fCycleTimeS 组态扫描周期
//           [秒]（限速积分基量）；② 覆盖 0.001~0.1 秒任务周期范围；
//           ③ 覆盖不到的区间由调用方按实际任务周期重设该引脚负责，
//           该假设挂编译验证债。同拍多窗配比约束（R100）：
//           tTrackTimeout > tShedHoldMin 不作要求（两窗职责独立：跟踪
//           失败窗对准伺服响应量级，卸荷保持窗对准雪滑落量级）。
// 开源溯源 (Origin)：道莅原创实现（参考跟踪支架雪载卸荷工程惯例 分类与参数域）
// 单位表：角度[度] / 角速度[度每秒] / 雪载[千克每平方米] / 阈值与回差
//         [千克每平方米] / 时间[ms] / 扫描周期[秒]
// 错误码表：16#0004_01E9 信息级（卸荷角到位提示，不置 bError）/
//           16#0004_01EA 信息级（复位角到位提示，不置 bError）/
//           16#0004_0309 故障级（组态非法：卸荷/复位角域、阈值/回差域、
//           限速/周期 <= 0 或任一输入非有限，置 bError）/ 16#0004_030A
//           故障级（角度反馈跟踪失败：反馈与命令偏差超容差持续超窗，
//           冻结命令安全侧，置 bError——该场景不可由 0309 的组态类
//           判据观测，属伺服跟踪独立域）/ 16#0004_030B 故障级兜底
//           （状态机落 ELSE，置 bError）
// 状态机：E_DL_SnowShedState（六态：eIdle=0 / eTrack=10 / eShedding=20 /
//           eShedHold=30 / eReturning=40 / eFault=99），CASE 含 ELSE
//           兜底，ELSE 置 030B 并冻结命令
// 边界行为：① 组态非法 → 故障态锁存，bReset 复位；② 限速逼近双向
//           适用（卸荷与复位均限速，防机构冲击）；③ 雪载回差防抖
//           （退出阈值 = 阈值 - 回差，阈值附近抖动防频动，R23 教训）；
//           ④ 卸荷保持最短时间未满不退出（防雪未滑落即回摆）；⑤ 故障
//           态命令冻结为最后合法值（跟踪失败时跳变比保持更危险）；
//           ⑥ 未使能命令冻结为 0 度并 bValid := FALSE。
// 修订历史：v1.0.0 2026-11-17 首版（R24 派单 · ROADMAP P1 §812）
//==============================================================================

(*------------------------------------------------------------------------------
 * 枚举: E_DL_SnowShedState（归属本功能块，同文件发布，全库唯一定义）
 * 含义: 雪载卸荷相位，每个成员在 CASE 中有且仅有一个标签。
 *-----------------------------------------------------------------------------*)
TYPE E_DL_SnowShedState :
(
    eIdle      := 0,   // 空闲：未使能 / Idle, not enabled
    eTrack     := 10,  // 跟踪：命令透传正常跟踪角 / Track, pass-through to the tracking angle
    eShedding  := 20,  // 卸荷中：限速逼近卸荷角 / Shedding, slewing to the shed angle
    eShedHold  := 30,  // 卸荷保持：最短保持计时 / Shed hold, minimum hold counting
    eReturning := 40,  // 复位中：限速逼近跟踪角 / Returning, slewing back to the tracking angle
    eFault     := 99   // 故障：组态非法/跟踪失败/非法状态 / Fault, config, tracking loss or illegal state
);
END_TYPE

FUNCTION_BLOCK FB_DL_TrackerSnowShedAngle
VAR_INPUT
    bEnable        : BOOL;                  // 卸荷控制使能 [—] / Shed control enable
    bReset         : BOOL;                  // 故障复位 [—]，上升沿清锁存 / Fault reset, rising edge clears latches
    bHeatSeason    : BOOL;                  // 采暖季窗有效 [—]（上层日历窗电平） / Heating-season window level
    fSnowLoadKgm2  : LREAL;                 // 雪载实测/估测 [千克每平方米] / Snow load [kg/m2]
    fTrackAngleDeg : LREAL;                 // 正常跟踪角 [度]（上层跟踪器透传） / Normal tracking angle [deg], pass-through
    fAngleFbDeg    : LREAL;                 // 角度反馈 [度] / Angle feedback [deg]
    fSnowThreshKgm2: LREAL := 5.0;          // 卸荷雪载阈 [千克每平方米]，须 > 0 / Shed threshold [kg/m2]
    fSnowHystKgm2  : LREAL := 1.0;          // 退出回差 [千克每平方米]，须 >= 0 且 < 阈值 / Exit hysteresis [kg/m2]
    fShedAngleDeg  : LREAL := 60.0;         // 卸荷角 [度]，域 [0, 90] / Shed angle [deg], domain 0..90
    fMaxSlewDegS   : LREAL := 2.0;          // 限速 [度每秒]，须 > 0 / Max slew rate [deg/s]
    fCycleTimeS    : LREAL := 0.01;         // 任务扫描周期 [秒]，须 > 0（R95 代理阈值） / Task scan cycle [s], must be > 0, R95 proxy
    tShedHoldMin   : TIME  := T#30S;        // 卸荷最短保持 [ms]，须 > 0 / Minimum shed hold [ms]
    fTrackTolDeg   : LREAL := 5.0;          // 反馈跟踪容差 [度]，须 > 0 / Feedback tracking tolerance [deg]
    tTrackTimeout  : TIME  := T#30S;        // 跟踪失败窗 [ms]，须 > 0 / Tracking-loss window [ms]
END_VAR
VAR_OUTPUT
    fAngleCmdDeg   : LREAL;                 // 角度命令 [度]（限速后，给驱动层） / Angle command [deg], post-slew
    bShedActive    : BOOL;                  // 卸荷活动 [—]（卸荷/保持态电平） / Shed active level
    eState         : E_DL_SnowShedState;    // 相位出口 [—] / Phase outlet
    eErr           : UDINT;                 // 错误码，0 = 无错，码位 16#0004_01E9 起信息级、16#0004_0309 起故障级（分带见错误码表） / Error code, 0 = no error, band info/fault per the code table
    bError         : BOOL;                  // 故障级标志，仅故障级错误置位 / Fault-class flag, set only on fault-level codes
    bValid         : BOOL;                  // 输出可用标志 / Outputs usable flag
END_VAR
VAR
    fbHold   : TON;                         // 卸荷保持计时（每拍无条件刷新）[ms] / Hold timer, refreshed unconditionally
    fbTrack  : TON;                         // 跟踪失败窗计时（每拍无条件刷新）[ms] / Tracking-loss timer, refreshed unconditionally
    _eState  : E_DL_SnowShedState := E_DL_SnowShedState.eIdle; // 当前相位 / Current phase
    _bCfgBad : BOOL;                        // 组态非法锁存 / Illegal config latch
    _bTrackBad: BOOL;                       // 跟踪失败锁存 / Tracking-loss latch
    _bInfoShed: BOOL;                       // 卸荷到位信息当拍标志 / Shed-arrival info flag of this scan
    _bInfoRet : BOOL;                       // 复位到位信息当拍标志 / Return-arrival info flag of this scan
    _fTarget  : LREAL;                      // 当前目标角 [度] / Current target angle [deg]
    _fStep    : LREAL;                      // 本拍限速步进 [度] / Per-scan slew step [deg]
    _bIllegal : BOOL;                       // 非法状态标志 / Illegal state flag
    _bInit    : BOOL := FALSE;              // 首扫标志，初值 FALSE 取非判定 / First-scan flag, tested negated
END_VAR
VAR CONSTANT
    DL_TSS_INF     : LREAL := 1.7976931348623157E308; // LREAL 幅值上限 / LREAL magnitude ceiling
    DL_TSS_EPS     : LREAL := 1.0E-6;       // 浮点判零/到位容差 [度] / Zero and arrival tolerance [deg]
    DL_TSS_SHED_MAX: LREAL := 90.0;         // 卸荷角域上限 [度] / Shed angle domain ceiling [deg]
    DL_TSS_ZERO    : LREAL := 0.0;          // 零值常量，避免裸字面量 [度] / Zero constant, avoids a bare literal
END_VAR

(*------------------------------------------------------------------------------
 * 段 1｜每拍预置：命令角保持语义（预置不清零，故障须冻结），标志预清零
 *      Command kept by design (frozen in fault), flags pre-cleared
 *-----------------------------------------------------------------------------*)
bShedActive := FALSE;                    // 卸荷电平先清（段 5 重置） / Shed level cleared first
eErr   := 16#0000_0000;                  // 错误码每拍重算 / Error code recomputed
bError := FALSE;                         // 故障标志每拍重算 / Fault flag recomputed
bValid := FALSE;                         // 可用标志每拍重算 / Usable flag recomputed
_bInfoShed := FALSE;                     // 卸荷信息预清零 / Shed info pre-cleared
_bInfoRet  := FALSE;                     // 复位信息预清零 / Return info pre-cleared
_bIllegal  := FALSE;                     // 非法状态预清零 / Illegal flag pre-cleared

(*------------------------------------------------------------------------------
 * 段 2｜首扫初始化
 *      First-scan initialisation
 *-----------------------------------------------------------------------------*)
IF NOT _bInit THEN
    _eState   := E_DL_SnowShedState.eIdle; // 相位空闲起步 / Phase starts idle
    _bCfgBad  := FALSE;                  // 组态锁存清零 / Config latch cleared
    _bTrackBad := FALSE;                 // 跟踪锁存清零 / Tracking latch cleared
    fAngleCmdDeg := DL_TSS_ZERO;         // 命令角从零起步 / Command starts at zero
    _bInit   := TRUE;                    // 首扫只做一次 / The first scan runs once
END_IF

(*------------------------------------------------------------------------------
 * 段 3｜组态防御闸：非有限（R79）+ 角度/阈值/限速/周期/时间窗域
 *      Configuration defense gates
 *-----------------------------------------------------------------------------*)
IF (fSnowLoadKgm2 <> fSnowLoadKgm2) OR (ABS(fSnowLoadKgm2) > DL_TSS_INF)
   OR (fTrackAngleDeg <> fTrackAngleDeg) OR (ABS(fTrackAngleDeg) > DL_TSS_INF)
   OR (fAngleFbDeg <> fAngleFbDeg) OR (ABS(fAngleFbDeg) > DL_TSS_INF)
   OR (fSnowThreshKgm2 <> fSnowThreshKgm2) OR (ABS(fSnowThreshKgm2) > DL_TSS_INF)
   OR (fSnowHystKgm2 <> fSnowHystKgm2) OR (ABS(fSnowHystKgm2) > DL_TSS_INF)
   OR (fShedAngleDeg <> fShedAngleDeg) OR (ABS(fShedAngleDeg) > DL_TSS_INF)
   OR (fMaxSlewDegS <> fMaxSlewDegS) OR (ABS(fMaxSlewDegS) > DL_TSS_INF)
   OR (fCycleTimeS <> fCycleTimeS) OR (ABS(fCycleTimeS) > DL_TSS_INF)
   OR (fTrackTolDeg <> fTrackTolDeg) OR (ABS(fTrackTolDeg) > DL_TSS_INF) THEN
    _bCfgBad := TRUE;                    // 非有限归组态非法锁存 / Non-finite folded into the config latch
END_IF
IF (NOT _bCfgBad) AND ((fSnowThreshKgm2 <= DL_TSS_EPS) OR (fSnowHystKgm2 < DL_TSS_ZERO)
   OR (fSnowHystKgm2 >= fSnowThreshKgm2) OR (fShedAngleDeg < DL_TSS_ZERO)
   OR (fShedAngleDeg > DL_TSS_SHED_MAX) OR (fMaxSlewDegS <= DL_TSS_EPS)
   OR (fCycleTimeS <= DL_TSS_EPS) OR (fTrackTolDeg <= DL_TSS_EPS)
   OR (tShedHoldMin <= T#0MS) OR (tTrackTimeout <= T#0MS)) THEN
    _bCfgBad := TRUE;                    // 角度/阈值/限速/周期/时间窗域非法锁存 / Angle, threshold, slew, cycle and window domains latched
END_IF
IF bReset THEN
    _bCfgBad   := FALSE;                 // 复位清组态锁存 / Reset clears the config latch
    _bTrackBad := FALSE;                 // 复位清跟踪锁存 / Reset clears the tracking latch
END_IF

(*------------------------------------------------------------------------------
 * 段 4｜双计时无条件刷新（R40：CASE 之外每拍必调）
 *      Two timers refreshed unconditionally per R40
 *-----------------------------------------------------------------------------*)
fbHold(IN := (_eState = E_DL_SnowShedState.eShedHold), PT := tShedHoldMin); // 卸荷保持窗 / Shed hold window
fbTrack(IN := (_eState = E_DL_SnowShedState.eShedding)
             OR (_eState = E_DL_SnowShedState.eReturning)
             OR (_eState = E_DL_SnowShedState.eTrack), PT := tTrackTimeout); // 跟踪失败窗（由段 5 IN 复判有效） / Tracking-loss window

(*------------------------------------------------------------------------------
 * 段 5｜相位机与限速逼近（CASE 含 ELSE 兜底；状态改写只出现在分支判据内，R39）
 *      Phase machine and the slew approach
 *-----------------------------------------------------------------------------*)
CASE _eState OF

    E_DL_SnowShedState.eIdle:              // 空闲：使能且组态合法进跟踪态
        IF bEnable AND (NOT _bCfgBad) THEN
            _eState := E_DL_SnowShedState.eTrack; // 进跟踪 / To track
        ELSIF bEnable AND _bCfgBad THEN
            _eState := E_DL_SnowShedState.eFault; // 组态非法进故障 / Illegal config to fault
        END_IF

    E_DL_SnowShedState.eTrack:             // 跟踪：透传正常角；采暖季且雪超阈进卸荷
        IF (NOT bEnable) OR _bCfgBad THEN
            _eState := E_DL_SnowShedState.eFault; // 异常转故障 / Anomaly, fault
        ELSE
            _fTarget := fTrackAngleDeg;    // 目标 = 正常跟踪角 / Target is the tracking angle
            IF bHeatSeason AND (fSnowLoadKgm2 > fSnowThreshKgm2) THEN
                _fTarget := fShedAngleDeg; // 目标切卸荷角 / Target switches to the shed angle
                _eState := E_DL_SnowShedState.eShedding; // 进卸荷 / To shedding
            END_IF
        END_IF

    E_DL_SnowShedState.eShedding:          // 卸荷：限速逼近；到位进保持；反馈失跟落故障
        IF (NOT bEnable) OR _bCfgBad THEN
            _eState := E_DL_SnowShedState.eFault; // 异常转故障 / Anomaly, fault
        ELSE
            _fTarget := fShedAngleDeg;     // 目标 = 卸荷角 / Target is the shed angle
            IF ABS(fAngleFbDeg - fAngleCmdDeg) > fTrackTolDeg THEN
                IF fbTrack.Q THEN
                    _bTrackBad := TRUE;    // 跟踪失败锁存（拍 N 进入） / Tracking loss latched
                    _eState := E_DL_SnowShedState.eFault; // 本拍转出：进故障冻结 / To fault, frozen
                END_IF
            ELSE
                _fTarget := fShedAngleDeg; // 到位判据仍按命令目标 / Arrival judged on the command target
                IF ABS(fAngleCmdDeg - _fTarget) <= DL_TSS_EPS THEN
                    _bInfoShed := TRUE;    // 卸荷角到位（信息级，拍 N 进入） / Shed angle reached, info
                    _eState := E_DL_SnowShedState.eShedHold; // 本拍转出：进保持 / To hold
                END_IF
            END_IF
        END_IF

    E_DL_SnowShedState.eShedHold:          // 保持：最短时间未满不退出；退出条件两判据 + 保持满
        IF (NOT bEnable) OR _bCfgBad THEN
            _eState := E_DL_SnowShedState.eFault; // 异常转故障 / Anomaly, fault
        ELSIF fbHold.Q AND (NOT bHeatSeason
               OR (fSnowLoadKgm2 < (fSnowThreshKgm2 - fSnowHystKgm2))) THEN
            _eState := E_DL_SnowShedState.eReturning; // 保持满且（季末或雪回差退出）进复位 / To returning
        END_IF

    E_DL_SnowShedState.eReturning:         // 复位：限速回跟踪角；到位进跟踪态
        IF (NOT bEnable) OR _bCfgBad THEN
            _eState := E_DL_SnowShedState.eFault; // 异常转故障 / Anomaly, fault
        ELSE
            _fTarget := fTrackAngleDeg;    // 目标 = 正常跟踪角 / Target is the tracking angle
            IF ABS(fAngleFbDeg - fAngleCmdDeg) > fTrackTolDeg THEN
                IF fbTrack.Q THEN
                    _bTrackBad := TRUE;    // 跟踪失败锁存 / Tracking loss latched
                    _eState := E_DL_SnowShedState.eFault; // 进故障冻结 / To fault, frozen
                END_IF
            ELSE
                IF ABS(fAngleCmdDeg - _fTarget) <= DL_TSS_EPS THEN
                    _bInfoRet := TRUE;     // 复位角到位（信息级） / Return angle reached, info
                    _eState := E_DL_SnowShedState.eTrack; // 进跟踪态 / To track
                END_IF
            END_IF
        END_IF

    E_DL_SnowShedState.eFault:             // 故障：复位沿且原因消失回跟踪态（命令保持冻结值）
        IF bReset AND (NOT _bCfgBad) AND (NOT _bTrackBad) THEN
            _eState := E_DL_SnowShedState.eTrack; // 回跟踪 / Back to track
        END_IF

    ELSE                                   // 非法状态兜底（R21：CASE 必带 ELSE）
        _bIllegal := TRUE;                 // 标记非法状态 / Flag the illegal state
        _eState := E_DL_SnowShedState.eFault; // 回故障态（命令冻结） / Back to fault, command frozen
END_CASE

(*------------------------------------------------------------------------------
 * 段 6｜限速逼近（跟踪/卸荷/复位态执行；故障/空闲冻结，不跳变）
 *      Slew approach in motion phases, frozen in fault and idle
 *-----------------------------------------------------------------------------*)
IF (_eState = E_DL_SnowShedState.eTrack)
   OR (_eState = E_DL_SnowShedState.eShedding)
   OR (_eState = E_DL_SnowShedState.eReturning)
   OR (_eState = E_DL_SnowShedState.eShedHold) THEN
    _fStep := fMaxSlewDegS * fCycleTimeS;  // 本拍限速步进 [度] / Per-scan slew step
    IF fAngleCmdDeg < (_fTarget - DL_TSS_EPS) THEN
        fAngleCmdDeg := MIN(fAngleCmdDeg + _fStep, _fTarget); // 上行限速逼近（饱和于目标） / Upward slew, saturated at the target
    ELSIF fAngleCmdDeg > (_fTarget + DL_TSS_EPS) THEN
        fAngleCmdDeg := MAX(fAngleCmdDeg - _fStep, _fTarget); // 下行限速逼近 / Downward slew
    END_IF
ELSIF _eState = E_DL_SnowShedState.eIdle THEN
    fAngleCmdDeg := DL_TSS_ZERO;           // 未使能命令归零（安全侧） / Not enabled, command to zero
END_IF
bShedActive := (_eState = E_DL_SnowShedState.eShedding)
            OR (_eState = E_DL_SnowShedState.eShedHold); // 卸荷活动电平挂状态量（R99） / Shed level bound to the states

(*------------------------------------------------------------------------------
 * 段 7｜码位出口与放行（故障级码 3 行内置 bError，R45/R101 配对）
 *      Code outlet and release, fault codes paired with bError
 *-----------------------------------------------------------------------------*)
IF _bIllegal THEN
    eErr   := 16#0004_030B;                // 故障级：状态机兜底 / Fault: state machine fallback
    bError := TRUE;                        // 置故障标志 / Raise the fault flag
ELSIF _bTrackBad THEN
    eErr   := 16#0004_030A;                // 故障级：角度反馈跟踪失败（命令冻结安全侧） / Fault: tracking loss, command frozen
    bError := TRUE;                        // 置故障标志 / Raise the fault flag
ELSIF _bCfgBad THEN
    eErr   := 16#0004_0309;                // 故障级：组态非法 / Fault: illegal configuration
    bError := TRUE;                        // 置故障标志 / Raise the fault flag
ELSIF _bInfoRet THEN
    eErr := 16#0004_01EA;                  // 信息级：复位角到位 / Info: return angle reached
ELSIF _bInfoShed THEN
    eErr := 16#0004_01E9;                  // 信息级：卸荷角到位 / Info: shed angle reached
END_IF

bValid := (NOT bError) AND bEnable AND (_eState <> E_DL_SnowShedState.eIdle); // 空闲/故障/未使能输出不可用 / Outputs unusable in idle, fault or disabled
eState := _eState;                       // 相位出口 / Phase outlet
END_FUNCTION_BLOCK

(* ---- FB_DL_TrapezoidProfilePlanner.st ---- *)
(*
  FB_DL_TrapezoidProfilePlanner —— 梯形/三角速度规划：起止速度不等，距离不足自动降级三角曲线，逐周期输出设定值与完成/超差标志
  分类：DL_Motion | 复杂度：4 | 轮次：R86
  开源溯源：道莅原创（clean-room 自研，纯 IEC 61131-3 通用算法），无外部代码引用
  许可证：MIT

  职责：按「目标位移 + 最大速度 + 最大加速度 + 起止速度 + 周期」做解析式梯形速度规划；
        当 fDa + fDd 超过目标位移时自动降级为三角曲线（峰值速度解含开方，负根 / 低于起止速度判规划失败）。
  输入契约：fDist 目标位移 [mm]（可为负，负号即反向）；fVelMax > 0；fAccMax > 0；
            fVelStart / fVelEnd 与 fDist 同号（按幅值参与规划）；fDt > 0 扫描周期 [s]。
  输出契约：fPosCmd / fVelCmd 为「相对起点的位移指令 / 速度指令」，符号随 fDist；
            xBusy 运动三相为 TRUE；xDone 到达终点的保持位；xOverrun 规划不可行或参数非法（锁存至下次启动沿）。
  边界：① 除零防护：fDt / fAccMax / fVelMax / fVp 全部前置判零；② 浮点比较一律用 DL_EPS 容差；
        ③ 起点段 eIdle 一次性解算全段时长，运动三相只做解析求值，无累积积分漂移；
        ④ 末拍精确落点（fPosCmd := fDist、fVelCmd := fVelEnd），消除解析式尾差；
        ⑤ 零全局耦合、零物理地址、零库件依赖（仅 SQRT / ABS 标准函数）。
*)

(*-----------------------------------------------------------------------------
 * 枚举: E_DL_TrapSeg（梯形规划段 / 状态，归属本文件，全库唯一定义）
 *----------------------------------------------------------------------------*)
TYPE E_DL_TrapSeg :
(
    eIdle   := 0,   // 空闲待启动 [—] / Idle, waiting for the start edge
    eAccel  := 1,   // 加速段（含三角曲线前半） [—] / Acceleration phase
    eCruise := 2,   // 匀速段（三角曲线时长为 0） [—] / Constant velocity phase
    eDecel  := 3,   // 减速段（含三角曲线后半） [—] / Deceleration phase
    eDone   := 4,   // 已到达终点（保持末值） [—] / Finished, outputs held
    eFault  := 5    // 规划失败 / 参数非法（锁存） [—] / Planning failed or invalid parameters
);
END_TYPE

FUNCTION_BLOCK FB_DL_TrapezoidProfilePlanner
VAR_INPUT
    xEnable   : BOOL  := TRUE;    // 使能，FALSE 时运动三相立即停机回空闲 [—] / Enable, false aborts motion to idle
    xStart    : BOOL  := FALSE;   // 启动（上升沿触发一次规划） [—] / Start, a rising edge triggers one plan
    fDist     : LREAL := 100.0;   // 目标位移，负值即反向 [mm] / Target displacement, negative means reverse
    fVelMax   : LREAL := 50.0;    // 最大允许速度（幅值） [mm/s] / Maximum allowed velocity magnitude
    fAccMax   : LREAL := 100.0;   // 最大允许加速度（幅值） [mm/s2] / Maximum allowed acceleration magnitude
    fVelStart : LREAL := 0.0;     // 起始速度（与 fDist 同号） [mm/s] / Start velocity, same sign as fDist
    fVelEnd   : LREAL := 0.0;     // 终止速度（与 fDist 同号） [mm/s] / End velocity, same sign as fDist
    fDt       : LREAL := 0.01;    // 扫描周期，必须 > 0 [s] / Scan period, must be positive
END_VAR
VAR_OUTPUT
    fPosCmd   : LREAL;                          // 位移指令（相对起点，带符号） [mm] / Position command relative to start
    fVelCmd   : LREAL;                          // 速度指令（带符号） [mm/s] / Velocity command with sign
    xBusy     : BOOL;                           // 运动进行中 [—] / Motion in progress
    xDone     : BOOL;                           // 已到达终点（保持位） [—] / Target reached, held
    xOverrun  : BOOL;                           // 规划不可行 / 参数非法（锁存） [—] / Planning overrun or invalid parameters
    xValid    : BOOL;                           // 本次规划有效 [—] / The current plan is valid
    eSeg      : E_DL_TrapSeg;                   // 当前段枚举 [—] / The active profile segment
END_VAR
VAR
    eState      : E_DL_TrapSeg;                 // 内部状态（与 eSeg 同步发布） [—] / Internal state mirrored to eSeg
    xStartPrev  : BOOL;                         // 启动信号上拍快照 [—] / Previous scan snapshot of xStart
    xEdgeStart  : BOOL;                         // 本拍启动上升沿 [—] / The start rising edge this scan
    xParamBad   : BOOL;                         // 参数 / 规划非法标志 [—] / Parameter or planning invalid flag
    xTriangle   : BOOL;                         // 三角曲线降级标志 [—] / Triangular profile degraded flag
    fSgn        : LREAL;                        // 位移方向符号（+1 / -1） [—] / Displacement direction sign
    fDistAbs    : LREAL;                        // 目标位移幅值 [mm] / Absolute target displacement
    fVStartAbs  : LREAL;                        // 起始速度幅值 [mm/s] / Absolute start velocity
    fVEndAbs    : LREAL;                        // 终止速度幅值 [mm/s] / Absolute end velocity
    fVp         : LREAL;                        // 实际峰值速度 [mm/s] / The effective peak velocity
    fVp2        : LREAL;                        // 峰值速度平方（开方前中间量） [mm2/s2] / Peak velocity squared
    fTa         : LREAL;                        // 加速段时长 [s] / Acceleration phase duration
    fTc         : LREAL;                        // 匀速段时长（三角曲线为 0） [s] / Cruise phase duration
    fTd         : LREAL;                        // 减速段时长 [s] / Deceleration phase duration
    fTtot       : LREAL;                        // 全段总时长 [s] / Total profile duration
    fDa         : LREAL;                        // 加速段位移 [mm] / Acceleration phase distance
    fDc         : LREAL;                        // 匀速段位移 [mm] / Cruise phase distance
    fDd         : LREAL;                        // 减速段位移 [mm] / Deceleration phase distance
    fTElapsed   : LREAL;                        // 已用时间 [s] / Elapsed time since the start edge
    fTd2        : LREAL;                        // 减速段内相对时间 [s] / Relative time inside the deceleration phase
    fS          : LREAL;                        // 位移幅值中间量 [mm] / Displacement magnitude intermediate
    fV          : LREAL;                        // 速度幅值中间量 [mm/s] / Velocity magnitude intermediate
END_VAR
VAR CONSTANT
    DL_EPS : LREAL := 1.0E-9;                   // 浮点比较容差 [—] / The floating point comparison tolerance
    DL_ZERO : LREAL := 0.0;                     // 浮点零常量 [—] / The floating point zero constant
    DL_TWO : LREAL := 2.0;                      // 浮点二常量 [—] / The floating point two constant
    DL_BIG : LREAL := 1.0E30;                   // 非有限值判据上界 [—] / The upper bound used to detect an infinite input
END_VAR

// 段 1｜周期无条件刷新：输出预置 + 启动沿提取（R7 无实例定时器，手工沿快照）
xEdgeStart := xStart AND NOT xStartPrev;        // 上升沿提取（上拍快照比对） / extract the rising edge
xDone := FALSE;                                 // 完成位预置假，CASE 内命中终点才置真 / preset done false
xBusy := FALSE;                                 // 忙碌位预置假，CASE 内运动三相置真 / preset busy false
xOverrun := FALSE;                              // 超差位预置假，CASE 内故障相置真 / preset overrun false
xValid := FALSE;                                // 规划有效位预置假，规划通过才置真 / preset valid false

// 段 2｜主状态机（ENUM + CASE，ELSE 拦截非法状态）
CASE eState OF

    E_DL_TrapSeg.eIdle:
        fPosCmd := DL_ZERO;                     // 空闲相位移指令归零 [mm] / idle position command zero
        fVelCmd := DL_ZERO;                     // 空闲相速度指令归零 [mm/s] / idle velocity command zero
        eSeg := E_DL_TrapSeg.eIdle;             // 段枚举发布空闲 / publish the idle segment
        IF xEdgeStart THEN                      // 收到启动沿 / a start edge arrived
            xParamBad := FALSE;                 // 参数闸标志复位 / reset the parameter gate flag
            fSgn := 1.0;                        // 方向符号预置正 / preset the sign positive
            IF fDist < DL_ZERO THEN             // 目标位移为负 / the target displacement is negative
                fSgn := -1.0;                   // 方向符号取负 / take the negative sign
            END_IF
            fDistAbs := ABS(fDist);             // 位移幅值 [mm] / the displacement magnitude
            fVStartAbs := ABS(fVelStart);       // 起始速度幅值 [mm/s] / the start velocity magnitude
            fVEndAbs := ABS(fVelEnd);           // 终止速度幅值 [mm/s] / the end velocity magnitude
            IF NOT xEnable THEN                 // 未使能启动 / started while disabled
                xParamBad := TRUE;              // 判参数非法 / mark the parameters invalid
            END_IF
            IF (fDist <> fDist) OR (fVelMax <> fVelMax) OR (fAccMax <> fAccMax)
               OR (fVelStart <> fVelStart) OR (fVelEnd <> fVelEnd) OR (fDt <> fDt)
               OR (ABS(fDist) > DL_BIG) OR (ABS(fVelMax) > DL_BIG) OR (ABS(fAccMax) > DL_BIG) THEN
                xParamBad := TRUE;              // 非有限值闸：NaN 或 Inf 一律判参数非法 / non-finite gate, NaN or Inf marks the parameters invalid
            END_IF
            IF fDt <= DL_ZERO THEN              // 周期非正（除零防护一） / the period is non positive
                xParamBad := TRUE;              // 判参数非法 / mark the parameters invalid
            END_IF
            IF fVelMax <= DL_ZERO THEN          // 最大速度非正（除零防护二） / the max velocity is non positive
                xParamBad := TRUE;              // 判参数非法 / mark the parameters invalid
            END_IF
            IF fAccMax <= DL_ZERO THEN          // 最大加速度非正（除零防护三） / the max acceleration is non positive
                xParamBad := TRUE;              // 判参数非法 / mark the parameters invalid
            END_IF
            IF fDistAbs <= DL_EPS THEN          // 目标位移近似为零 / the target displacement is near zero
                xParamBad := TRUE;              // 判参数非法 / mark the parameters invalid
            END_IF
            IF fVStartAbs > fVelMax + DL_EPS THEN // 起始速度越最大速度 / the start velocity above the maximum
                xParamBad := TRUE;              // 判参数非法 / mark the parameters invalid
            END_IF
            IF fVEndAbs > fVelMax + DL_EPS THEN // 终止速度越最大速度 / the end velocity above the maximum
                xParamBad := TRUE;              // 判参数非法 / mark the parameters invalid
            END_IF
            IF (fVelStart * fVelEnd) < -DL_EPS THEN // 起止速度异号，需过零，本件不支持 / opposite signs unsupported
                xParamBad := TRUE;              // 判参数非法 / mark the parameters invalid
            END_IF
            IF NOT xParamBad THEN               // 参数全通过才做规划 / plan only when all parameters pass
                fDa := (fVelMax * fVelMax - fVStartAbs * fVStartAbs) / (DL_TWO * fAccMax); // 满速加速段位移 [mm]
                fDd := (fVelMax * fVelMax - fVEndAbs * fVEndAbs) / (DL_TWO * fAccMax);     // 满速减速段位移 [mm]
                IF (fDa + fDd) <= fDistAbs THEN // 位移足够走梯形 / enough distance for a trapezoid
                    xTriangle := FALSE;         // 梯形标志 / trapezoidal profile
                    fVp := fVelMax;             // 峰值速度取最大速度 [mm/s] / the peak equals the maximum
                    fDc := fDistAbs - fDa - fDd;// 匀速段位移 [mm] / the cruise distance
                ELSE                            // 位移不足，降级三角曲线 / degrade to a triangle
                    xTriangle := TRUE;          // 三角标志 / triangular profile
                    fVp2 := (DL_TWO * fAccMax * fDistAbs + fVStartAbs * fVStartAbs + fVEndAbs * fVEndAbs) / DL_TWO; // 峰值速度平方 [mm2/s2]
                    IF fVp2 <= DL_ZERO THEN // 负根或零根，距离不足以起停 / negative root, distance too short
                        xParamBad := TRUE;  // 判规划失败 / mark the planning failure
                    ELSE
                        fVp := SQRT(fVp2);  // 峰值速度取正根 [mm/s] / take the positive root
                        IF (fVp < fVStartAbs - DL_EPS) OR (fVp < fVEndAbs - DL_EPS) THEN // 峰值低于起止速度，距离连加速都装不下
                            xParamBad := TRUE;  // 判规划失败 / mark the planning failure
                        END_IF
                    END_IF
                    IF NOT xParamBad THEN       // 三角曲线重算各段位移 / recompute the triangle distances
                        fDa := (fVp * fVp - fVStartAbs * fVStartAbs) / (DL_TWO * fAccMax); // 加速段位移 [mm]
                        fDd := (fVp * fVp - fVEndAbs * fVEndAbs) / (DL_TWO * fAccMax);     // 减速段位移 [mm]
                        fDc := DL_ZERO;     // 三角曲线无匀速段 [mm] / no cruise distance in a triangle
                    END_IF
                END_IF
            END_IF
            IF NOT xParamBad THEN               // 位移段解算通过后解时长 / solve the phase durations
                fTa := (fVp - fVStartAbs) / fAccMax; // 加速段时长 [s] / the acceleration duration
                fTd := (fVp - fVEndAbs) / fAccMax;   // 减速段时长 [s] / the deceleration duration
                IF fVp > DL_EPS THEN            // 峰值速度非零（除零防护四） / the peak velocity is positive
                    fTc := fDc / fVp;           // 匀速段时长 [s] / the cruise duration
                ELSE
                    fTc := DL_ZERO;             // 零速退化，匀速段记零 [s] / degenerate, cruise duration zero
                END_IF
                fTtot := fTa + fTc + fTd;       // 全段总时长 [s] / the total duration
                IF fTtot <= DL_EPS THEN         // 总时长为零，规划不可行 / the total duration is zero
                    xParamBad := TRUE;          // 判规划失败 / mark the planning failure
                END_IF
            END_IF
            IF xParamBad THEN                   // 任一闸判失败 / any gate failed
                eState := E_DL_TrapSeg.eFault;  // 迁入故障相（锁存） / enter the fault state, latched
                eSeg := E_DL_TrapSeg.eFault;    // 段枚举发布故障 / publish the fault segment
                fPosCmd := DL_ZERO;             // 位移指令归零 [mm] / position command zero
                fVelCmd := DL_ZERO;             // 速度指令归零 [mm/s] / velocity command zero
                xOverrun := TRUE;               // 置超差位 [—] / raise the overrun flag
            ELSE                                // 规划通过 / the plan passes
                fTElapsed := DL_ZERO;           // 已用时间清零 [s] / clear the elapsed time
                xValid := TRUE;                 // 置规划有效 [—] / raise the valid flag
                xBusy := TRUE;                  // 置忙碌位 [—] / raise the busy flag
                fPosCmd := DL_ZERO;             // 起点位移指令为零 [mm] / the start position command
                fVelCmd := fVelStart;           // 起点速度指令为起始速度 [mm/s] / the start velocity command
                eSeg := E_DL_TrapSeg.eAccel;    // 段枚举发布加速段 / publish the acceleration segment
                eState := E_DL_TrapSeg.eAccel;  // 迁入加速段 / enter the acceleration phase
            END_IF
        END_IF

    E_DL_TrapSeg.eAccel, E_DL_TrapSeg.eCruise, E_DL_TrapSeg.eDecel:
        IF NOT xEnable THEN                     // 使能撤销，立即停机 / the enable dropped, stop at once
            eState := E_DL_TrapSeg.eIdle;       // 回空闲相 / back to idle
            eSeg := E_DL_TrapSeg.eIdle;         // 段枚举发布空闲 / publish the idle segment
            fVelCmd := DL_ZERO;                 // 速度指令归零 [mm/s] / velocity command zero
            fPosCmd := DL_ZERO;                 // 位移指令归零 [mm] / position command zero
        ELSE
            fTElapsed := fTElapsed + fDt;       // 累加已用时间 [s]（fDt > 0 已在规划闸证明）
            IF fTElapsed <= fTa THEN            // 落在加速段时间窗内 / inside the acceleration window
                fS := fVStartAbs * fTElapsed + 0.5 * fAccMax * fTElapsed * fTElapsed; // 位移幅值 [mm]
                fV := fVStartAbs + fAccMax * fTElapsed;                              // 速度幅值 [mm/s]
                eSeg := E_DL_TrapSeg.eAccel;    // 段枚举发布加速段 / publish the acceleration segment
            ELSIF fTElapsed <= (fTa + fTc) THEN // 落在匀速段时间窗内 / inside the cruise window
                fS := fDa + fVp * (fTElapsed - fTa); // 位移幅值 [mm] / the displacement magnitude
                fV := fVp;                      // 速度幅值取峰值 [mm/s] / the velocity magnitude equals the peak
                eSeg := E_DL_TrapSeg.eCruise;   // 段枚举发布匀速段 / publish the cruise segment
            ELSE                                // 落在减速段时间窗内 / inside the deceleration window
                fTd2 := fTElapsed - fTa - fTc;  // 减速段内相对时间 [s] / the relative time inside deceleration
                fS := fDa + fDc + fVp * fTd2 - 0.5 * fAccMax * fTd2 * fTd2; // 位移幅值 [mm]
                fV := fVp - fAccMax * fTd2;     // 速度幅值 [mm/s] / the velocity magnitude
                eSeg := E_DL_TrapSeg.eDecel;    // 段枚举发布减速段 / publish the deceleration segment
            END_IF
            IF fS > fDistAbs THEN               // 位移幅值上越界钳位 / clamp the displacement magnitude
                fS := fDistAbs;                 // 钳到目标位移 [mm] / clamp to the target
            END_IF
            IF fS < DL_ZERO THEN                // 位移幅值下越界钳位 / clamp the lower side
                fS := DL_ZERO;                  // 钳到零 [mm] / clamp to zero
            END_IF
            IF fV < DL_ZERO THEN                // 速度幅值下越界钳位 / clamp the velocity magnitude
                fV := DL_ZERO;                  // 钳到零 [mm/s] / clamp to zero
            END_IF
            fPosCmd := fSgn * fS;               // 带符号位移指令出口 [mm] / the signed position command
            fVelCmd := fSgn * fV;               // 带符号速度指令出口 [mm/s] / the signed velocity command
            xBusy := TRUE;                      // 运动三相置忙碌 [—] / raise busy during the motion phases
            xValid := TRUE;                     // 运动三相规划仍有效 [—] / the plan stays valid while moving
            IF fTElapsed >= (fTtot - DL_EPS) THEN // 到达总时长 / the total duration is reached
                fPosCmd := fDist;               // 末拍精确落点 [mm] / the exact final position
                fVelCmd := fVelEnd;             // 末拍精确末速 [mm/s] / the exact final velocity
                xDone := TRUE;                  // 置完成位 [—] / raise the done flag
                xBusy := FALSE;                 // 撤忙碌位 [—] / drop the busy flag
                eSeg := E_DL_TrapSeg.eDone;     // 段枚举发布完成 / publish the done segment
                eState := E_DL_TrapSeg.eDone;   // 迁入完成相（锁存末值） / enter the done state, outputs held
            END_IF
        END_IF

    E_DL_TrapSeg.eDone:
        fPosCmd := fDist;                       // 保持精确终点 [mm] / hold the exact final position
        fVelCmd := fVelEnd;                     // 保持精确末速 [mm/s] / hold the exact final velocity
        xDone := TRUE;                          // 保持完成位 [—] / hold the done flag
        xValid := TRUE;                         // 保持规划有效 [—] / hold the valid flag
        eSeg := E_DL_TrapSeg.eDone;             // 保持段枚举完成 / hold the done segment
        IF xEdgeStart THEN                      // 完成后再启动一次 / restarted from the done state
            eState := E_DL_TrapSeg.eIdle;       // 回空闲相，下一拍重新规划 / back to idle for a fresh plan
        END_IF

    E_DL_TrapSeg.eFault:
        fPosCmd := DL_ZERO;                     // 故障相位移指令归零 [mm] / fault state position zero
        fVelCmd := DL_ZERO;                     // 故障相速度指令归零 [mm/s] / fault state velocity zero
        xOverrun := TRUE;                       // 故障锁存回放超差位 [—] / replay the latched overrun flag
        eSeg := E_DL_TrapSeg.eFault;            // 段枚举发布故障 / publish the fault segment
        IF (NOT xStart) AND NOT xEnable THEN    // 撤启动信号且使能撤销 / start released and enable dropped
            eState := E_DL_TrapSeg.eIdle;       // 唯一解除路径：该条件沿回空闲 / the only clear edge back to idle
        END_IF

ELSE
    eState := E_DL_TrapSeg.eFault;              // 非法枚举值一律拦入故障相 / trap any illegal state value
    eSeg := E_DL_TrapSeg.eFault;                // 段枚举发布故障 / publish the fault segment
    fPosCmd := DL_ZERO;                         // 位移指令归零 [mm] / position command zero
    fVelCmd := DL_ZERO;                         // 速度指令归零 [mm/s] / velocity command zero
    xOverrun := TRUE;                           // 置超差位 [—] / raise the overrun flag
END_CASE

// 段 3｜启动信号上拍快照（位于主体末尾，保证本拍沿检测用的是上拍值）
xStartPrev := xStart;                           // 末尾刷新上拍快照 / refresh the previous snapshot at the end
END_FUNCTION_BLOCK

(* ---- FB_DL_TurretToolSelect.st ---- *)
(*
  ==================================================================
  组件名 Component  : FB_DL_TurretToolSelect
  分类   Category   : DL_Motion
  前缀   Naming     : FB_DL_ ｜ b/n/u/f/t/e/st 类型前缀制（R265）
  复杂度 Complexity  : 高
  版本   Version    : 1.0.1
  功能   Purpose    : 刀塔就近方向换刀选择（刀位环计数 + 最短路径 + 当前刀位校验状态机）。
  来源   Source     : t1-6-plcopen（PLCopen 刀塔换刀公开语义）
  平台   Platform   : 纯 IEC 61131-3（R_TRIG / CASE / MOD），三平台通用
  分工声明 Split     : 与 FB_DL_TurretIndexSeq（顺序换刀属主，若在册）分工——本件
                      只做就近方向解算与校验，不做顺序全环巡检（R216 双向互引）。
  作者   Author     : 道莅代码库 · PLC 编程专家（R61）
  归属 Ownership     : E_DL_TurretPhase 属主为本文件（全库唯一定义，R264）；
                      引用件只引用不重声明。
  ------------------------------------------------------------------
  边界 Boundary     :
                      一 刀位号域闸 [1, n] 钳位：越域钳位后仍以钳位值解算（信息级
                         08A6），不拒单（换刀请求尽量满足）；
                      二 就近方向判据整数进位点自证：环差 diff = (req − cur) MOD n，
                         恰对径（diff·2 = n）两向量等长时写死取正向（CW），判据
                         全整数精确比较，无浮点；
                      三 换刀指令单拍脉冲 bToolChange（R256 统一出口预置）；
                      四 状态机 CASE 必带 ELSE 兜底；R_TRIG 段 0 无条件刷新（R7）；
                      五 故障锁存解除式自证：刀位数组态非法（<1 或 >24）锁存
                         08A7，bReset 上升沿解除（恒可达，R152 自证）；
                      七 故障相迁入完备（v1.0.1 修 D3）：段 4 之后设统一迁入闸
                         （_bFault 且当前相 ≠ eFault 即迁 eFault），eMoving 的故障
                         出口亦直接迁 eFault，eFault 成为可达相而非死相位；
                      八 不删 eFault 相的理由（诊断保真）：eFault 是 R274 要求的
                         状态机完整性成员，且与 FB_DL_SingleAxis 族故障相命名一致；
                         删相会让「组态非法」与「空闲」在 eState 出口上不可分，
                         现场读 eState=eIdle 且 bError=TRUE 时无法区分「未换刀」
                         与「组态故障」，损失诊断保真；
                      六 无全局、无外部变量、无物理地址。
  错误码   Codes    :
    16#0004_08A6【信息级】刀位号或刀位数越域已钳位（[1, 24]）
    16#0004_08A7【故障级】刀位数组态非法（<1 或 >24），锁存至复位沿
  验收   Acceptance :
    算法已证（脚本）：未跑 ｜ 编译器已证（三平台）：未跑
    V1 n=8、cur=1、req=3 → 正向 2 步；V2 cur=1、req=7 → 反向 2 步
    V3 n=8、cur=1、req=5（对径）→ 正向 4 步（进位点写死取正）
    V4 req=0 → 钳到 1、码 08A6；n=0 → 码 08A7 锁存
    V5 组态非法（uToolCnt=0）→ eState=eFault 且 bError=TRUE 同拍（v1.0.1 回归向量）
    V6 故障态下 bReset 上升沿且组态已合法 → 清锁存、迁 eIdle
    V7 正常换刀全程 → eState 轨迹 eIdle→eMoving→eIdle，eFault 不出现
  修订记录 Revision  :
    2026-11-21  v1.0.0  R61 首版（批 4 · 序号 15）
    2026-11-21  v1.0.1  R62-D3 返修：①段 4 后加故障统一迁入闸（R274 迁入完备性），补 eFault 死相位；②eMoving 的 ELSIF _bFault 出口由 eIdle 改为 eFault；③eFault 出口「NOT _bFault 才迁出」保持不变；④不删相理由（诊断保真）写入头注释。注：盘面实测入库版本为 v1.0.0（计划书假设 R61 已发 v1.0.1），按实测优先、禁跳号递增一次至 v1.0.1
  ==================================================================
*)
TYPE E_DL_TurretPhase :
(
    eIdle   := 0,  // 空闲：等换刀指令沿 / idle, waiting for the change edge
    eMoving := 10, // 换刀进行：等到位反馈 / moving, waiting for the in position feedback
    eFault  := 20  // 故障：组态非法，锁存待复位 / fault, the illegal configuration latched
);
END_TYPE

FUNCTION_BLOCK FB_DL_TurretToolSelect
VAR_INPUT
    bExec     : BOOL := FALSE;  // 换刀指令电平，上升沿解算并发单拍 / the change command level
    bInPos    : BOOL := FALSE;  // 刀塔到位反馈电平 [-] / the turret in position feedback
    bReset    : BOOL := FALSE;  // 故障复位电平，上升沿清锁存 / the fault reset level
    uCurTool  : UDINT := 1;     // 当前刀位号 [刀位]，域 [1, 24] / the current tool number
    uReqTool  : UDINT := 1;     // 请求刀位号 [刀位]，域 [1, 24] / the requested tool number
    uToolCnt  : UDINT := 8;     // 刀位总数 [刀位]，合法域 1..24 / the tool count, legal from one to twenty four
END_VAR
VAR_OUTPUT
    bDirCW      : BOOL := FALSE;          // 方向指示：TRUE 正向（CW）[-] / the direction indicator, true for the forward
    uSteps      : UDINT := 0;             // 换刀步数 [步] / the change step count
    bToolChange : BOOL := FALSE;          // 换刀指令单拍脉冲 [-] / the change command one shot pulse
    bDone       : BOOL := FALSE;          // 换刀完成单拍脉冲 [-] / the change done one shot pulse
    eState      : E_DL_TurretPhase;       // 主状态机当前态 [状态] / the current state
    bError      : BOOL := FALSE;          // 故障锁存位（与锁存同源，R191）/ the fault bit from the latch
    bValid      : BOOL := FALSE;          // 解算可用标志 [-] / the solve usable flag
    eErr        : UDINT := 16#0000_0000;  // 错误码，0 = 正常 / the error code, zero is ok
END_VAR
VAR
    _bInit    : BOOL := FALSE;                        // 首拍初始化标志（R310）/ the first scan flag
    _eState   : E_DL_TurretPhase := E_DL_TurretPhase.eIdle; // 内部状态寄存器 / the internal state register
    _bFault   : BOOL := FALSE;                        // 组态故障锁存副本（仅复位沿清除）/ the fault latch copy
    _nCur     : DINT := 1;                            // 钳位后当前刀位 [刀位] / the clamped current tool
    _nReq     : DINT := 1;                            // 钳位后请求刀位 [刀位] / the clamped requested tool
    _nCnt     : DINT := 8;                            // 钳位后刀位数 [刀位] / the clamped tool count
    _nDiff    : DINT := 0;                            // 环差 [步] / the ring difference
    _nSteps   : DINT := 0;                            // 步数工作副本 [步] / the step count copy
    _bCW      : BOOL := FALSE;                        // 方向工作副本 / the direction copy
    _bChange  : BOOL := FALSE;                        // 换刀单拍内部位，段 1 预清段 5 映射 / the internal change bit
    _bDone    : BOOL := FALSE;                        // 完成单拍内部位 / the internal done bit
    _bClamp   : BOOL := FALSE;                        // 钳位标记（逐拍重算）/ the clamp flag recomputed
    rtExec    : R_TRIG; // 换刀指令沿实例，段 0 无条件刷新 / the command edge instance
    rtReset   : R_TRIG; // 复位沿实例，段 0 无条件刷新 / the reset edge instance
END_VAR
VAR CONSTANT
    DL_TTS_NMAX : DINT := 24; // 刀位容量上界 [刀位] / the tool capacity bound
END_VAR

// 段 0｜沿检测无条件周期刷新（禁入分支，R7）/ segment 0, the unconditional refresh
rtExec(CLK := bExec); // 换刀指令沿 / the command edge
rtReset(CLK := bReset); // 复位沿 / the reset edge

// 段 1｜首拍初始化与单拍标志预清（R310 / FB32-1 / R256）/ segment 1, the first scan init and the preset
IF NOT _bInit THEN // 首拍一拍 / the first scan
    _bInit := TRUE; // 置首拍标志 / raise the first scan flag
    _bFault := FALSE; // 故障锁存显式清零 / clear the fault latch explicitly
    _eState := E_DL_TurretPhase.eIdle; // 状态显式落空闲 / place the state to idle
END_IF
IF rtReset.Q THEN // 复位沿（作用域：清锁存 + 迁相位，R311 声明）/ the reset edge with the declared scope
    _bFault := FALSE; // 清锁存（解除路径：复位沿恒可达，R152 自证）/ clear the latch
    _eState := E_DL_TurretPhase.eIdle; // 迁回空闲 / back to idle
END_IF
_bChange := FALSE; // 换刀单拍预清零 / preset the change bit false
_bDone := FALSE; // 完成单拍预清零 / preset the done bit false
_bClamp := FALSE; // 钳位标记预清零 / preset the clamp flag false

// 段 2｜域闸与钳位（整数全精确，边界一二五）/ segment 2, the domain gate with the clamps
_nCnt := UDINT_TO_DINT(uToolCnt); // 刀位数升位接管 / take the tool count widened
IF (_nCnt < 1) OR (_nCnt > DL_TTS_NMAX) THEN // 刀位数组态非法（0807 → 08A7 独立码）/ the illegal tool count
    _bFault := TRUE; // 锁存故障（08A7）/ latch the fault
END_IF
IF _nCnt < 1 THEN // 下界钳位（防环运算除零取模）/ the floor clamp guarding the modulo
    _nCnt := 1; // 钳到一 / clamp to one
END_IF
IF _nCnt > DL_TTS_NMAX THEN // 上界钳位 / the ceiling clamp
    _nCnt := DL_TTS_NMAX; // 钳到容量 / clamp to the capacity
END_IF
_nCur := UDINT_TO_DINT(uCurTool); // 当前刀位接管 / take the current tool
_nReq := UDINT_TO_DINT(uReqTool); // 请求刀位接管 / take the requested tool
IF (_nCur < 1) OR (_nCur > _nCnt) OR (_nReq < 1) OR (_nReq > _nCnt) THEN // 刀位号越域（信息级钳位，边界一）/ the tool numbers out of the domain
    _bClamp := TRUE; // 置钳位标记 / raise the clamp flag
END_IF
IF _nCur < 1 THEN // 当前刀位下界钳位 / the current floor clamp
    _nCur := 1; // 钳到一 / clamp to one
END_IF
IF _nCur > _nCnt THEN // 当前刀位上界钳位 / the current ceiling clamp
    _nCur := _nCnt; // 钳到总数 / clamp to the count
END_IF
IF _nReq < 1 THEN // 请求刀位下界钳位 / the requested floor clamp
    _nReq := 1; // 钳到一 / clamp to one
END_IF
IF _nReq > _nCnt THEN // 请求刀位上界钳位 / the requested ceiling clamp
    _nReq := _nCnt; // 钳到总数 / clamp to the count
END_IF

// 段 3｜就近方向解算（全整数精确比较，进位点写死取正向，边界二）/ segment 3, the nearest direction solve in exact integers
_nDiff := ((_nReq - _nCur) MOD _nCnt + _nCnt) MOD _nCnt; // 环差归一到 [0, n-1]（双 MOD 防负数取模方言差异）/ the ring difference normalized
IF _nDiff = 0 THEN // 同刀位：零步 / the same tool, zero steps
    _nSteps := 0; // 零步 / zero steps
    _bCW := TRUE; // 零步时方向寄存器按正向表态（无方向语义）/ the direction placeholder forward
ELSIF (_nDiff * 2) = _nCnt THEN // 恰对径（进位点）：两向等长，写死取正向（边界二）/ the diametric point takes the forward by the declared rule
    _nSteps := _nDiff; // 正向步数 / the forward steps
    _bCW := TRUE; // 正向 / forward
ELSIF (_nDiff * 2) < _nCnt THEN // 正向更近 / the forward is nearer
    _nSteps := _nDiff; // 正向步数 / the forward steps
    _bCW := TRUE; // 正向 / forward
ELSE // 反向更近 / the reverse is nearer
    _nSteps := _nCnt - _nDiff; // 反向步数 / the reverse steps
    _bCW := FALSE; // 反向 / reverse
END_IF

// 段 4｜主状态机（ENUM + CASE，ELSE 兜底；指令沿消费带全量闸位复检，R274）/ segment 4, the main machine
CASE _eState OF
    E_DL_TurretPhase.eIdle: // 空闲相 / the idle phase
        IF rtExec.Q AND (NOT _bFault) THEN // 指令沿 + 闸位复检（R274）/ the command edge with the gate recheck
            IF _nSteps = 0 THEN // 同刀位校验：直接完成（整数精确比较，边界二）/ the same tool verified by the exact integer compare
                _bDone := TRUE; // 置完成单拍 / raise the done bit
            ELSE // 异刀位：发换刀单拍并迁入移动相 / a different tool, raise the change pulse and enter moving
                _bChange := TRUE; // 置换刀单拍 / raise the change bit
                _eState := E_DL_TurretPhase.eMoving; // 迁入移动相 / enter the moving phase
            END_IF
        END_IF
    E_DL_TurretPhase.eMoving: // 移动相：等到位反馈 / the moving phase
        IF bInPos THEN // 到位反馈（同刀位目标校验后完成）/ the in position feedback
            _bDone := TRUE; // 置完成单拍 / raise the done bit
            _eState := E_DL_TurretPhase.eIdle; // 迁回空闲 / back to idle
        ELSIF _bFault THEN // 前置条件消失出口（直接迁故障相，不经 eIdle，v1.0.1 修 D3）/ the prerequisite gone exit straight to the fault phase
            _eState := E_DL_TurretPhase.eFault; // 迁入故障相（与统一迁入闸同向，避免同拍先迁 idle 再被拉回）/ enter the fault phase, aligned with the unified gate
        END_IF
    E_DL_TurretPhase.eFault: // 故障相：等复位沿（解除可达，边界五）/ the fault phase until the reset
        IF NOT _bFault THEN // 锁存已清才迁出 / the exit after the latch cleared
            _eState := E_DL_TurretPhase.eIdle; // 迁回空闲 / back to idle
        END_IF
    ELSE // 非法枚举值拦截 / the illegal enumeration guard
        _eState := E_DL_TurretPhase.eIdle; // 落回空闲 / force back to idle
        _bFault := TRUE; // 置锁存 / latch the fault
END_CASE

// 段 4b｜故障统一迁入闸（置于状态机之后、解除段之外，R274 迁入完备性；v1.0.1 修 D3）/ segment 4b, the unified fault entry gate
IF _bFault AND (_eState <> E_DL_TurretPhase.eFault) THEN // 已锁存但当前不在故障相（含 eIdle 检出与非法枚举值兜底）/ latched but not yet in the fault phase
    _eState := E_DL_TurretPhase.eFault; // 任何相检出故障一律落故障相，eFault 由此可达 / any phase with a latch lands in the fault phase, which makes it reachable
END_IF

// 段 5｜统一出口（内部副本单点映射；故障码锁存回放，R187）/ segment 5, the unified outlet
bDirCW := _bCW; // 方向出口 / the direction outlet
uSteps := DINT_TO_UDINT(_nSteps); // 步数出口（值已证非负）/ the step outlet proven non negative
bToolChange := _bChange; // 换刀单拍出口 / the change pulse outlet
bDone := _bDone; // 完成单拍出口 / the done pulse outlet
eState := _eState; // 状态出口 / the state outlet
bError := _bFault; // 故障位出口（与锁存同源）/ the fault bit outlet
bValid := NOT _bFault; // 解算可用标志 / the solve usable flag
IF _bFault THEN // 故障锁存回放（R187）/ the latched fault replays
    eErr := 16#0004_08A7; // 故障级：刀位数组态非法 / fault grade, the illegal tool count
ELSIF _bClamp THEN // 钳位（信息级不置 bError，R285）/ the clamp informational
    eErr := 16#0004_08A6; // 信息级：刀位号越域已钳位 / informational, the tool numbers clamped
ELSE // 无事件 / no event
    eErr := 16#0000_0000; // 正常 / ok
END_IF
END_FUNCTION_BLOCK
